(* IEC 61131-3 sources: daoli-st-library/DL_Algo (part 10) *)

(* ---- FB_DL_CoolingTowerApproachCalc.st ---- *)
//==============================================================================
// 功能块：FB_DL_CoolingTowerApproachCalc ｜ 中文名称：冷却塔逼近度计算与风机台数优化建议
// 所属子库：DL_Algo ｜ 版本：v1.0.0 ｜ 兼容：CODESYS V3.5+ / TwinCAT 3 / 汇川 InoProShop
// 功能描述：逼近度 = 冷却水出水温度 − 湿球温度（湿球由
//           FC_DL_WetBulbTempCalc v1.1.0 计算，组合调用不内联）；逼近度
//           滑动均值（1~60 拍窗）进入目标带判断；带外给出增/减风机台数
//           建议（单拍脉冲），带内保持。优化纪律：逼近度优先、N+1 冗余
//           （减台不低于 1 台）、换台最小间隔（tMinStageTime，被阻延沿
//           发一次 3402 提示）、湿球贴物理极限逼近度时加机无益（禁止
//           建议加机）。只出建议，不直接控风机（启停时序由上位轮值件
//           裁决，本件零执行输出）。
// 开源溯源 (Origin)：道莅原创实现（参考 公开工程惯例 分类与参数域）
// 单位表：温度[摄氏度] / 相对湿度[%] / 大气压[Pa] / 逼近度[K] / 台数[台] / 换台间隔[min] / 均值窗[拍]
// 错误码表：16#0002_3401 信息级（逼近度小于 0，出水低于湿球，传感器可疑，
//           不给任何换台建议，不置 bError）/ 16#0002_3402 信息级（换台
//           请求被最小间隔阻延，阻延沿发一次，不置 bError）/
//           16#0002_3405 预留禁用（不得挪用）/ 16#0002_3410 故障级（台
//           数或算法组态非法，置 bError）/ 16#0002_3411 故障级（输入非
//           有限或湿球件故障透传，置 bError）/ 16#0002_3412 预留禁用
//           （不得挪用）
// 状态机：E_DL_ApproachState（eIdle=0 / eWarmup=10 / eMonitor=20 /
//           eStageUpPending=30 / eStageDownPending=40 / eFault=99），
//           CASE 含 ELSE 兜底，ELSE 复用 3411（§3 未为本件单列兜底槽，
//           不得越段加码）并回 eFault、脉冲全撤、建议保持（安全侧）
// 边界行为：① 湿球件 bError 或 bValid 为假 → 透传为故障 3411 +
//           bWetBulbFault，锁存型标志只在故障相处置（R115），下游信息级
//           码（钳位提示）不升格；② fApproachK 小于 0（热力学不可能，
//           传感器可疑）→ 信息 3401 + bValid := FALSE + 不给任何换台
//           建议，可疑样本不入均值窗（防污染统计）；③ nFanRunning 大于
//           nFanTotal 或 nFanTotal 小于 1 或均值窗/目标/带宽组态非法 →
//           故障 3410；④ 浮点输入非有限 → 故障 3411；⑤ 换台请求受
//           tMinStageTime 约束，被阻延 → 信息 3402（阻延沿发一次，不每
//           拍刷），阻延期间挂 eStageUpPending/eStageDownPending，退出
//           条件两条：间隔到且需求仍在（发请求回 eMonitor）或带偏差
//           消失/需求翻转（不发请求回 eMonitor）；⑥ 湿球贴物理极限逼
//           近度（常量 2.0 K）且台数已满 → bNoFurtherGain，禁止建议加
//           机；首次换台请求不受守卫约束（上电无历史换台）；⑦ 失能 →
//           建议台数保持、脉冲全撤、bValid := FALSE；⑧ 恢复首拍窗口
//           清空重走暖机；守卫定时器经请求签发「断输入一拍」重启计时
//           （R40 家族）；⑨ 上电首拍 bValid := FALSE。
// 修订历史：v1.0.0 2026-11-17 首版（R25 派单 · §4.3）
//==============================================================================
(*------------------------------------------------------------------------------
 * 枚举: E_DL_ApproachState（归属 DL_Algo，与 FB_DL_CoolingTowerApproachCalc 同文件）
 *----------------------------------------------------------------------------*)
TYPE E_DL_ApproachState :
(
    eIdle             := 0,   // 失能/待机：建议保持，脉冲全撤 / Idle: suggestion held, pulses withdrawn
    eWarmup           := 10,  // 暖机：均值窗未满，只观测不出建议 / Warmup: window not full, observe only
    eMonitor          := 20,  // 监视：带内保持或按需即时发换台请求 / Monitor: hold in band or issue request at once
    eStageUpPending   := 30,  // 增台请求被最小间隔阻延，等守卫计时 / Increase request blocked by min interval
    eStageDownPending := 40,  // 减台请求被最小间隔阻延，等守卫计时 / Decrease request blocked by min interval
    eFault            := 99   // 故障兜底态：组态非法/非有限/下游透传 / Fault fallback
);
END_TYPE
FUNCTION_BLOCK FB_DL_CoolingTowerApproachCalc
VAR_INPUT
    fCondOutC        : LREAL;                  // 冷却水出水温度 [摄氏度] / Condenser water outlet temperature [degC]
    fAmbDryC         : LREAL;                  // 环境干球温度 [摄氏度] / Ambient dry-bulb temperature [degC]
    fRhPct           : LREAL;                  // 环境相对湿度 [百分数] / Ambient relative humidity [percent]
    fPressPa         : LREAL := 101325.0;      // 大气压 [Pa]，引脚注入非魔法数 / Atmospheric pressure [Pa], pin-injected
    nFanTotal        : INT;                    // 可投风机台数 [台]，1~8 / Total available fans, 1~8
    nFanRunning      : INT;                    // 当前运行台数 [台]，0~8 / Currently running fans, 0~8
    fApproachTargetK : LREAL := 4.0;           // 目标逼近度 [K] / Target approach [K]
    fApproachTolK    : LREAL := 0.5;           // 逼近度带宽半宽 [K] / Approach band half-width [K]
    tMinStageTime    : TIME := T#5M;           // 换台最小间隔 [min] / Minimum interval between stage changes [min]
    nWinSamples      : INT := 10;              // 均值窗长度 [拍]，1~60 / Moving-average window length, 1~60
    bEnable          : BOOL;                   // 总使能 / Master enable
    bReset           : BOOL;                   // 复位，上升沿清状态与窗口 / Reset, rising edge clears state and window
END_VAR
VAR_OUTPUT
    fWetBulbC        : LREAL;                  // 湿球温度 [摄氏度]，下游件输出透传 / Wet-bulb temperature [degC], passed through
    fApproachK       : LREAL;                  // 即时逼近度 [K]，出水减湿球 / Instantaneous approach [K]
    fApproachAvgK    : LREAL;                  // 逼近度滑动均值 [K] / Moving-average approach [K]
    nFanCmd          : INT;                    // 建议运行台数 [台]，失能保持 / Suggested running fans, held on disable
    bIncReq          : BOOL;                   // 增台建议，单拍脉冲 / Increase suggestion, one-scan pulse
    bDecReq          : BOOL;                   // 减台建议，单拍脉冲 / Decrease suggestion, one-scan pulse
    bNoFurtherGain   : BOOL;                   // 湿球已贴物理极限逼近度，加机无益 / Wet bulb at physical floor, more fans useless
    bWetBulbFault    : BOOL;                   // 湿球下游件故障透传标志，只在故障相处置 / Wet-bulb downstream fault pass-through flag
    eErr             : UDINT;                  // 错误码，0 = 无错，码位 16#0002_3401 起信息级、16#0002_3410 起故障级（分带见错误码表） / Error code, 0 = no error, band info/fault per the code table
    bError           : BOOL;                   // 故障级标志，仅故障级错误置位 / Fault-class flag, set only on fault-level codes
    bValid           : BOOL;                   // 建议数据可用标志，失能/故障闸显式 FALSE / Suggestion usable flag, explicit FALSE on disable/fault gates
    eState           : E_DL_ApproachState;     // 主状态机当前状态 / Current state of the main state machine
END_VAR
VAR
    fWbOut           : LREAL;                  // 湿球件输出暂存 [摄氏度] / Wet-bulb output staging [degC]
    bWbClamped       : BOOL;                   // 湿球件钳位标志透传 / Wet-bulb clamped flag pass-through
    eWbErr           : UDINT;                  // 湿球件错误码暂存 / Wet-bulb error code staging
    bWbErr           : BOOL;                   // 湿球件故障标志暂存 / Wet-bulb fault flag staging
    bWbOk            : BOOL;                   // 湿球件可用且无故障 / Wet-bulb usable and fault-free
    fbReset          : R_TRIG;                 // 复位上升沿检测实例 / Reset rising edge detector
    fbBlockTrig      : R_TRIG;                 // 换台阻延上升沿检测实例（3402 一次触发）/ Stage-block rising edge detector, 3402 once per edge
    fbStageGuard     : TON;                    // 换台最小间隔守卫定时器 / Stage interval guard timer
    bGuardKick       : BOOL;                   // 守卫定时器断输入一拍标志（R40 家族）/ Guard timer one-scan kick flag
    afWinBuf         : ARRAY[0..59] OF LREAL;  // 逼近度滑动窗缓冲 [K] / Approach sliding window buffer [K]
    nWinIdx          : INT;                    // 窗写指针 [—] / Window write pointer
    uWinFill         : UDINT;                  // 窗已填充数 [拍] / Window filled count
    fWinSum          : LREAL;                  // 窗内累加和 [K]，增量维护 / Window running sum [K], incrementally maintained
    fApproachNew     : LREAL;                  // 本拍新逼近度样本 [K] / New approach sample this scan [K]
    bBadSensor       : BOOL;                   // 逼近度小于 0，传感器可疑 / Approach negative, sensor suspect
    bNeedInc         : BOOL;                   // 本拍需要增台（实时重算）/ Increase needed this scan, recomputed
    bNeedDec         : BOOL;                   // 本拍需要减台（实时重算）/ Decrease needed this scan, recomputed
    bGuardOk         : BOOL;                   // 守卫放行：无历史换台或间隔已满 / Guard released: no history or interval elapsed
    bBlockedNow      : BOOL;                   // 本拍换台请求被阻延 / Stage request blocked this scan
    bStageEverReq    : BOOL;                   // 激活以来是否签发过换台请求 / Any stage request issued since activation
    bFanCmdInit      : BOOL;                   // 建议台数是否已初始化 / Suggestion count initialized flag
    bActiveCalc      : BOOL;                   // 本拍处于可计算状态（暖机/监视/阻延挂起）/ Computable state this scan
END_VAR
VAR CONSTANT
    DL_CTWR_CODE_INFO_1 : UDINT := 16#0002_3401;   // 信息级槽 1（逼近度小于 0） / info slot 1
    DL_CTWR_CODE_INFO_2 : UDINT := 16#0002_3402;   // 信息级槽 2（换台请求被阻延） / info slot 2
    DL_CTWR_CODE_RSV_1  : UDINT := 16#0002_3405;   // 预留禁用（不得挪用） / reserved, do not use
    DL_CTWR_CODE_FLT_1  : UDINT := 16#0002_3410;   // 故障级槽 1（台数或组态非法） / fault slot 1
    DL_CTWR_CODE_FLT_2  : UDINT := 16#0002_3411;   // 故障级槽 2（非有限或湿球透传） / fault slot 2
    DL_CTWR_CODE_RSV_2  : UDINT := 16#0002_3412;   // 预留禁用（不得挪用） / reserved, do not use
    DL_AP_ZERO       : LREAL := 0.0;           // 零值常量，避免裸字面量 [—] / Zero constant, avoids a bare literal
    DL_AP_INF        : LREAL := 1.7976931348623157E308;  // LREAL 幅值上限，Inf 判据 / LREAL magnitude ceiling, Inf criterion
    DL_AP_TOL        : LREAL := 1.0E-6;        // 浮点比较容差 [—] / Float comparison tolerance
    DL_AP_WIN_MAX    : INT   := 60;            // 均值窗长度上限 [拍] / Moving-average window ceiling
    DL_AP_FAN_MAX    : INT   := 8;             // 风机台数上限 [台] / Fan count ceiling
    DL_AP_FAN_MIN    : INT   := 1;             // N+1 冗余最低运行台数 [台] / Minimum running fans for N+1 redundancy
    DL_AP_PHYS_FLOOR : LREAL := 2.0;           // 物理极限逼近度 [K]，贴限判加机无益 / Physical floor approach [K], gain-limit criterion
END_VAR

(*------------------------------------------------------------------------------
 * 段 1｜无条件刷新区（红线 5）：沿检测与守卫定时器在任何分支之外周期调用
 *----------------------------------------------------------------------------*)
fbReset(CLK := bReset);                        // 复位沿检测无条件刷新 / reset edge refreshed unconditionally
fbStageGuard(IN := bEnable AND NOT bGuardKick, // 断输入一拍重启计时（R40 家族）/ break input one scan to restart timing
             PT := tMinStageTime);             // 守卫门槛 = 换台最小间隔 / guard threshold = min stage interval
bGuardKick := FALSE;                           // kick 标志单拍自清（本拍签发请求时由状态机重置位）/ kick flag self-clears, state machine re-sets on issue

(*------------------------------------------------------------------------------
 * 段 2｜复位沿处理（改写置于沿后，防吞沿 R39）
 *----------------------------------------------------------------------------*)
IF fbReset.Q THEN
    eState        := E_DL_ApproachState.eIdle;
    eErr          := 16#0000_0000;             // 复位清码 / reset clears code
    bError        := FALSE;                    // 复位清故障 / reset clears fault
    uWinFill      := 0;                        // 窗口清空重走暖机 / window cleared, warmup again
    nWinIdx       := 0;                        // 写指针归零 / write pointer zeroed
    fWinSum       := DL_AP_ZERO;               // 累加和清零 / sum zeroed
    fApproachAvgK := DL_AP_ZERO;               // 均值出口清零 / average output zeroed
    bIncReq       := FALSE;                    // 脉冲全撤 / pulses withdrawn
    bDecReq       := FALSE;                    // 脉冲全撤 / pulses withdrawn
    bNoFurtherGain := FALSE;                   // 贴限标志清除 / gain-limit flag cleared
    bBadSensor    := FALSE;                    // 传感器可疑标志清除 / suspect flag cleared
    bStageEverReq := FALSE;                    // 换台历史清零，首个请求放行 / stage history cleared, first request released
    bFanCmdInit   := FALSE;                    // 建议台数待重初始化 / suggestion count re-initialized
END_IF

(*------------------------------------------------------------------------------
 * 段 3｜非有限输入闸（浮点引脚逐个：NaN 自反判 + Inf 幅值上限判，R79）
 *----------------------------------------------------------------------------*)
IF (fCondOutC <> fCondOutC) OR (ABS(fCondOutC) >= DL_AP_INF)
   OR (fAmbDryC <> fAmbDryC) OR (ABS(fAmbDryC) >= DL_AP_INF)
   OR (fRhPct <> fRhPct) OR (ABS(fRhPct) >= DL_AP_INF)
   OR (fPressPa <> fPressPa) OR (ABS(fPressPa) >= DL_AP_INF)
   OR (fApproachTargetK <> fApproachTargetK) OR (ABS(fApproachTargetK) >= DL_AP_INF)
   OR (fApproachTolK <> fApproachTolK) OR (ABS(fApproachTolK) >= DL_AP_INF) THEN
    eState := E_DL_ApproachState.eFault;
    eErr   := DL_CTWR_CODE_FLT_2;                  // 故障级：输入非有限 / fault: non-finite input
    bError := TRUE;                            // 故障级必置 bError（R45 配对）/ fault-class pairs with bError
    bValid := FALSE;                           // 输出不可用 / outputs unusable
    bIncReq := FALSE;                          // 脉冲全撤安全侧 / pulses withdrawn, safe side
    bDecReq := FALSE;                          // 脉冲全撤安全侧 / pulses withdrawn, safe side
    bNoFurtherGain := FALSE;                   // 故障态不判贴限 / gain-limit not judged in fault
    RETURN;
END_IF

(*------------------------------------------------------------------------------
 * 段 4｜组态合法性闸（台数域/主从关系/窗长/目标/带宽）
 *----------------------------------------------------------------------------*)
IF (nFanTotal < DL_AP_FAN_MIN) OR (nFanTotal > DL_AP_FAN_MAX)
   OR (nFanRunning < 0) OR (nFanRunning > nFanTotal)
   OR (nWinSamples < 1) OR (nWinSamples > DL_AP_WIN_MAX)
   OR (fApproachTargetK <= DL_AP_TOL) OR (fApproachTolK <= DL_AP_TOL) THEN
    eState := E_DL_ApproachState.eFault;
    eErr   := DL_CTWR_CODE_FLT_1;                  // 故障级：台数或算法组态非法 / fault: fan or algorithm config invalid
    bError := TRUE;                            // 故障级必置 bError（R45 配对）/ fault-class pairs with bError
    bValid := FALSE;                           // 输出不可用 / outputs unusable
    bIncReq := FALSE;                          // 脉冲全撤安全侧 / pulses withdrawn, safe side
    bDecReq := FALSE;                          // 脉冲全撤安全侧 / pulses withdrawn, safe side
    bNoFurtherGain := FALSE;                   // 故障态不判贴限 / gain-limit not judged in fault
    RETURN;
END_IF

(*------------------------------------------------------------------------------
 * 段 5｜湿球组合调用：每拍恰好一次，不内联不复制（R115 透传纪律）
 *----------------------------------------------------------------------------*)
FC_DL_WetBulbTempCalc(fTempC := fAmbDryC, fRh := fRhPct, fPress := fPressPa,
                      fWetBulbC => fWbOut, bClamped => bWbClamped,
                      eErr => eWbErr, bError => bWbErr, bValid => bWbOk);
fWetBulbC := fWbOut;                           // 湿球出口透传 / wet-bulb output pass-through
IF bWbErr OR (NOT bWbOk) THEN
    bWetBulbFault := TRUE;                     // 下游故障透传标志 / downstream fault pass-through flag
ELSE
    bWetBulbFault := FALSE;                    // 下游正常，信息级钳位不升格 / downstream ok, info-level clamp not escalated
END_IF

(*------------------------------------------------------------------------------
 * 段 6｜逼近度计算与滑动窗维护（仅在使能、湿球可用、传感器不可疑时推进）
 *----------------------------------------------------------------------------*)
bActiveCalc := bEnable AND (NOT bWetBulbFault)
           AND (eState = E_DL_ApproachState.eWarmup
             OR eState = E_DL_ApproachState.eMonitor
             OR eState = E_DL_ApproachState.eStageUpPending
             OR eState = E_DL_ApproachState.eStageDownPending);  // 可计算状态判据 / computable-state predicate
bBadSensor := FALSE;                           // 传感器可疑标志逐拍重判 / suspect flag re-judged per scan
IF bActiveCalc THEN
    fApproachK := fCondOutC - fWetBulbC;       // 即时逼近度 = 出水 − 湿球 [K] / instantaneous approach = outlet minus wet bulb
    bBadSensor := fApproachK < -DL_AP_TOL;     // 热力学不可能，传感器可疑 / thermodynamically impossible, sensor suspect
    IF bBadSensor THEN
        // 可疑样本不入窗，均值保持（防污染统计）/ suspect sample not pushed, average held
    ELSE
        IF uWinFill < INT_TO_UDINT(nWinSamples) THEN
            uWinFill := uWinFill + 1;          // 窗未满：填充数递增 / window not full: fill count up
            fWinSum := fWinSum + fApproachK;   // 累加和并入新样本 / sum absorbs new sample
            afWinBuf[nWinIdx] := fApproachK;   // 写入当前槽 / write current slot
        ELSE
            fWinSum := fWinSum - afWinBuf[nWinIdx] + fApproachK;  // 窗满：换出旧值并入新值 / window full: swap out old, absorb new
            afWinBuf[nWinIdx] := fApproachK;   // 覆盖当前槽 / overwrite current slot
        END_IF
        nWinIdx := (nWinIdx + 1) MOD nWinSamples;  // 写指针环形推进，nWinSamples 已闸大于 0 / ring-advance write pointer, divisor gated
        fApproachAvgK := fWinSum / UDINT_TO_LREAL(uWinFill);  // 均值 = 和/填充数，填充数已闸大于 0 / average, fill count gated
    END_IF
END_IF

(*------------------------------------------------------------------------------
 * 段 7｜决策块：带偏差实时重算（阻延挂起态也用同一决策，需求翻转即退出）
 *----------------------------------------------------------------------------*)
bNeedInc := FALSE;                             // 增台需求逐拍重判 / increase need re-judged per scan
bNeedDec := FALSE;                             // 减台需求逐拍重判 / decrease need re-judged per scan
bNoFurtherGain := FALSE;                       // 贴限标志逐拍重判，非计算态不残留 / gain-limit flag re-judged per scan
bGuardOk := (NOT bStageEverReq) OR fbStageGuard.Q;  // 守卫放行：无历史换台或最小间隔已满 / guard released
IF bActiveCalc AND (NOT bBadSensor) THEN
    IF NOT bFanCmdInit THEN
        nFanCmd := nFanRunning;                // 建议台数首拍初始化为当前运行台数 / suggestion initialized to running count
        bFanCmdInit := TRUE;                   // 初始化完成 / initialization done
    END_IF
    bNoFurtherGain := (fApproachK <= DL_AP_PHYS_FLOOR) AND (nFanRunning >= nFanTotal);  // 贴物理极限且台数已满，加机无益 / at physical floor with all fans on
    IF (fApproachAvgK - fApproachTargetK) > fApproachTolK THEN
        bNeedInc := (nFanRunning < nFanTotal) AND (NOT bNoFurtherGain);  // 偏热且有余量：增台 / too hot with headroom: increase
    ELSIF (fApproachTargetK - fApproachAvgK) > fApproachTolK THEN
        bNeedDec := (nFanRunning > DL_AP_FAN_MIN);  // 偏冷且高于冗余下限：减台 / too cold above redundancy floor: decrease
    END_IF
END_IF

(*------------------------------------------------------------------------------
 * 段 8｜阻延沿检测（无条件周期调用，CLK 为本拍阻延判据，3402 沿发一次）
 *----------------------------------------------------------------------------*)
bBlockedNow := bActiveCalc AND (NOT bBadSensor) AND (bNeedInc OR bNeedDec) AND (NOT bGuardOk);  // 本拍阻延判据 / blocked predicate this scan
fbBlockTrig(CLK := bBlockedNow);               // 阻延沿检测无条件刷新 / block edge refreshed unconditionally

(*------------------------------------------------------------------------------
 * 段 9｜状态机：CASE 含 ELSE 兜底。bIncReq/bDecReq 为单拍脉冲：本段开头
 *       先无条件撤脉冲，状态机内按需重置位（先撤后置，不跨拍残留）。
 *----------------------------------------------------------------------------*)
bIncReq := FALSE;                              // 单拍脉冲先撤 / one-scan pulse withdrawn first
bDecReq := FALSE;                              // 单拍脉冲先撤 / one-scan pulse withdrawn first

CASE eState OF

    E_DL_ApproachState.eIdle:
        bValid := FALSE;                       // 失能闸显式不可用（R72）/ explicit FALSE on disable gate
        eErr := 16#0000_0000;                  // 待机无错 / no error in idle
        bError := FALSE;                       // 待机无故障 / no fault in idle
        bWetBulbFault := FALSE;                // 待机不透传故障相（R115：只在故障相处置）/ pass-through only in fault phase
        bNoFurtherGain := FALSE;               // 待机不判贴限 / gain-limit not judged in idle
        IF bEnable THEN
            IF bWetBulbFault THEN
                eState := E_DL_ApproachState.eFault;   // 湿球不可用直接进故障 / unusable wet bulb enters fault
                eErr := DL_CTWR_CODE_FLT_2;    // 故障级：湿球件故障透传 / fault: wet-bulb pass-through
                bError := TRUE;                // 故障级必置 bError / fault-class pairs with bError
            ELSE
                eState := E_DL_ApproachState.eWarmup;  // 使能且湿球可用进暖机 / enable with valid wet bulb enters warmup
            END_IF
        END_IF

    E_DL_ApproachState.eWarmup:
        eErr := 16#0000_0000;                  // 暖机默认无错 / warmup defaults to no error
        bError := FALSE;                       // 暖机默认无故障 / warmup defaults to no fault
        bValid := FALSE;                       // 暖机期窗口未满不可用 / unusable during warmup
        IF NOT bEnable THEN
            eState := E_DL_ApproachState.eIdle;        // 失能回待机 / disable returns to idle
        ELSIF bWetBulbFault THEN
            eState := E_DL_ApproachState.eFault;       // 下游故障进故障态 / downstream fault enters fault state
            eErr := DL_CTWR_CODE_FLT_2;        // 故障级：湿球件故障透传 / fault: wet-bulb pass-through
            bError := TRUE;                    // 故障级必置 bError / fault-class pairs with bError
        ELSIF bBadSensor THEN
            eErr := DL_CTWR_CODE_INFO_1;       // 信息级：逼近度小于 0，传感器可疑 / info: negative approach, sensor suspect
            bValid := FALSE;                   // 传感器可疑，不给建议 / suspect sensor, no advice
        ELSIF uWinFill >= INT_TO_UDINT(nWinSamples) THEN
            eState := E_DL_ApproachState.eMonitor;     // 均值窗已满进监视 / window full enters monitor
        END_IF

    E_DL_ApproachState.eMonitor:
        IF NOT bEnable THEN
            eState := E_DL_ApproachState.eIdle;        // 失能回待机 / disable returns to idle
            bValid := FALSE;                   // 失能闸显式不可用（R72）/ explicit FALSE on disable gate
        ELSIF bWetBulbFault THEN
            eState := E_DL_ApproachState.eFault;
            eErr := DL_CTWR_CODE_FLT_2;        // 故障级：湿球件故障透传 / fault: wet-bulb pass-through
            bError := TRUE;                    // 故障级必置 bError / fault-class pairs with bError
            bValid := FALSE;                   // 故障闸显式不可用 / explicit FALSE on fault gate
        ELSIF bBadSensor THEN
            eErr := DL_CTWR_CODE_INFO_1;       // 信息级：逼近度小于 0 / info: negative approach
            bError := FALSE;                   // 信息级不置 bError / info never raises bError
            bValid := FALSE;                   // 传感器可疑，不给建议（边界行为②）/ suspect sensor, no advice
        ELSE
            eErr := 16#0000_0000;              // 正常监视清码 / normal monitor clears code
            bError := FALSE;                   // 正常监视清故障 / normal monitor clears fault
            bValid := TRUE;                    // 建议数据可用 / suggestion usable
            IF bNeedInc OR bNeedDec THEN
                IF bGuardOk THEN
                    IF bNeedInc THEN
                        bIncReq := TRUE;       // 增台建议单拍脉冲 / increase pulse
                        nFanCmd := nFanRunning + 1;    // 建议台数加一 / suggested count up
                    ELSE
                        bDecReq := TRUE;       // 减台建议单拍脉冲 / decrease pulse
                        nFanCmd := nFanRunning - 1;    // 建议台数减一 / suggested count down
                    END_IF
                    bStageEverReq := TRUE;     // 记录换台历史 / record stage history
                    bGuardKick := TRUE;        // 守卫定时器断输入一拍重启 / guard timer kicked one scan
                ELSE
                    IF bNeedInc THEN
                        eState := E_DL_ApproachState.eStageUpPending;  // 增台请求被阻延挂起 / increase request blocked, pending
                    ELSE
                        eState := E_DL_ApproachState.eStageDownPending;  // 减台请求被阻延挂起 / decrease request blocked, pending
                    END_IF
                END_IF
            END_IF
        END_IF

    E_DL_ApproachState.eStageUpPending:
        IF NOT bEnable THEN
            eState := E_DL_ApproachState.eIdle;
            bValid := FALSE;                   // 失能闸显式不可用（R72）/ explicit FALSE on disable gate
        ELSIF bWetBulbFault THEN
            eState := E_DL_ApproachState.eFault;
            eErr := DL_CTWR_CODE_FLT_2;
            bError := TRUE;
            bValid := FALSE;
        ELSIF bBadSensor THEN
            eState := E_DL_ApproachState.eMonitor;     // 传感器可疑，需求作废回监视 / suspect sensor, need voided, back to monitor
            eErr := DL_CTWR_CODE_INFO_1;
            bError := FALSE;
            bValid := FALSE;
        ELSIF NOT bNeedInc THEN
            eState := E_DL_ApproachState.eMonitor;     // 需求消失退出（第二条退出条件）/ need vanished, second exit condition
            eErr := 16#0000_0000;              // 回监视清码 / clear code on return
            bValid := TRUE;                    // 回监视数据可用 / usable on return
        ELSIF fbStageGuard.Q THEN
            bIncReq := TRUE;                   // 间隔到且需求仍在：签发增台 / interval elapsed with need: issue increase
            nFanCmd := nFanRunning + 1;        // 建议台数加一 / suggested count up
            bStageEverReq := TRUE;             // 记录换台历史 / record stage history
            bGuardKick := TRUE;                // 守卫定时器断输入一拍重启 / guard timer kicked one scan
            eState := E_DL_ApproachState.eMonitor;     // 签发后回监视 / back to monitor after issue
            eErr := 16#0000_0000;              // 阻延解除清码 / clear code on release
            bValid := TRUE;                    // 数据可用 / usable
        ELSE
            bValid := TRUE;                    // 挂起期间建议数据仍可用 / suggestion usable while pending
        END_IF

    E_DL_ApproachState.eStageDownPending:
        IF NOT bEnable THEN
            eState := E_DL_ApproachState.eIdle;
            bValid := FALSE;                   // 失能闸显式不可用（R72）/ explicit FALSE on disable gate
        ELSIF bWetBulbFault THEN
            eState := E_DL_ApproachState.eFault;
            eErr := DL_CTWR_CODE_FLT_2;
            bError := TRUE;
            bValid := FALSE;
        ELSIF bBadSensor THEN
            eState := E_DL_ApproachState.eMonitor;     // 传感器可疑，需求作废回监视 / suspect sensor, need voided, back to monitor
            eErr := DL_CTWR_CODE_INFO_1;
            bError := FALSE;
            bValid := FALSE;
        ELSIF NOT bNeedDec THEN
            eState := E_DL_ApproachState.eMonitor;     // 需求消失退出（第二条退出条件）/ need vanished, second exit condition
            eErr := 16#0000_0000;              // 回监视清码 / clear code on return
            bValid := TRUE;                    // 回监视数据可用 / usable on return
        ELSIF fbStageGuard.Q THEN
            bDecReq := TRUE;                   // 间隔到且需求仍在：签发减台 / interval elapsed with need: issue decrease
            nFanCmd := nFanRunning - 1;        // 建议台数减一 / suggested count down
            bStageEverReq := TRUE;             // 记录换台历史 / record stage history
            bGuardKick := TRUE;                // 守卫定时器断输入一拍重启 / guard timer kicked one scan
            eState := E_DL_ApproachState.eMonitor;     // 签发后回监视 / back to monitor after issue
            eErr := 16#0000_0000;              // 阻延解除清码 / clear code on release
            bValid := TRUE;                    // 数据可用 / usable
        ELSE
            bValid := TRUE;                    // 挂起期间建议数据仍可用 / suggestion usable while pending
        END_IF

    ELSE
        eState := E_DL_ApproachState.eFault;   // 非法状态兜底 / illegal-state fallback
        eErr   := DL_CTWR_CODE_FLT_2;          // 兜底复用故障级槽 2（§3 未单列兜底槽，不得越段加码）/ fallback reuses fault slot 2
        bError := TRUE;                        // 故障级必置 bError / fault-class pairs with bError
        bValid := FALSE;                       // 输出不可用 / outputs unusable
        bIncReq := FALSE;                      // 脉冲全撤安全侧 / pulses withdrawn, safe side
        bDecReq := FALSE;                      // 脉冲全撤安全侧 / pulses withdrawn, safe side
END_CASE

(*------------------------------------------------------------------------------
 * 段 10｜信息级收口：阻延沿发一次 3402（不每拍刷，见边界行为⑤）
 *----------------------------------------------------------------------------*)
IF fbBlockTrig.Q THEN
    eErr := DL_CTWR_CODE_INFO_2;               // 信息级：换台请求被最小间隔阻延 / info: stage request blocked by interval
    bError := FALSE;                           // 信息级不置 bError / info never raises bError
END_IF
END_FUNCTION_BLOCK

(* ---- FB_DL_CoolingTowerOpt.st ---- *)
(*
  Component : FB_DL_CoolingTowerOpt
  Category  : DL_Algo
  Type      : FB
  Version   : 1.0.0
  CodeSeg   : 16#02_3_5F
  Summary   : 冷却塔群控逼近度优化：湿球逼近度控制律 + 塔群投切决策（最小开机数 + 防震荡死区）。
              Cooling tower approach optimization: wet-bulb approach control law plus staging with min-on units and deadband.
  溯源声明  : 道莅自研 clean-room
  边界安全  : 温度/台数非有限（NaN 自反 + Inf 上限）拦截；塔数域闸（1..8，防数组越界）；
              最小开机数域闸（1..nTowers，防全停）与投切错峰窗（自复位 TON）防频繁投切；
              投切决策带对称死区（防震荡）；风机设定值输出过 RateLimiter 限速；
              全浮点比较带 fEps 容差；计数防回卷。
  复用      : 无
*)

FUNCTION_BLOCK FB_DL_CoolingTowerOpt
VAR_INPUT
    bRun          : BOOL;              (* 优化使能 · Enable *)
    fWetBulbC     : LREAL;             (* 湿球温度 [degC] · Wet-bulb temperature *)
    fOutTC        : LREAL;             (* 塔群出水温度 [degC] · Tower outlet temperature *)
    fApprTargetC  : LREAL := 3.0;      (* 逼近度目标 [K] · Approach target *)
    fDeadK        : LREAL := 0.5;      (* 投切死区 [K]，防震荡 · Staging deadband *)
    nTowersAvail  : INT   := 4;        (* 可用塔数 [台]，域 1 到 8 · Available towers *)
    nMinOn        : INT   := 1;        (* 最小开机数 [台] · Minimum on units *)
    tStaggerMs    : TIME  := T#30000MS; (* 投切错峰窗 [ms] · Stagger window *)
    fFanStepPct   : LREAL := 2.0;      (* 风机设定每拍最大步进 [％] · Fan setpoint max step *)
    fEps          : LREAL := 1.0E-6;   (* 浮点判零容差 [实数域] · Floating zero tolerance *)
END_VAR
VAR_OUTPUT
    aTowerCmd : ARRAY[1..8] OF BOOL;    (* 各塔投切指令 [引脚] · Per-tower commands *)
    nRunCnt   : INT;                    (* 当前开机数 [台] · Currently running count *)
    fApprNowC : LREAL;                  (* 当前逼近度 [K] · Current approach *)
    fFanSetPct: LREAL;                  (* 风机群设定值输出 [％]，已限速 · Rate-limited fan setpoint *)
    bError    : BOOL;                   (* 故障标志，与故障码配对 · Fault flag paired with codes *)
    uErrorId  : UDINT;                  (* 事件码 16#0000_005F，0 无事件 · Event code *)
END_VAR
VAR
    _eState   : (eStHold := 0, eStAdd := 1, eStDrop := 2);  (* 内部决策状态 / Internal decision state *)
    uCode     : WORD;    (* 码位暂存，每拍重算 [码] · Code staging *)
    tonStagger: TON;     (* 投切错峰窗 [ms]，自复位振荡 · Stagger timer, self-reset *)
    bSigOk    : BOOL;    (* 输入有效标志 · Input validity flag *)
    bTick     : BOOL;    (* 错峰窗到点脉冲 [脉冲] · Stagger tick pulse *)
    nI        : INT;     (* 塔循环下标 [索引] · Tower loop index *)
    fFanTgt   : LREAL;   (* 风机设定目标 [％] · Fan setpoint target *)
    fStep     : LREAL;   (* 本拍设定步进 [％] · Actual step this scan *)
    nCycles   : UDINT;   (* 有效拍计数 [拍]，防回卷 · Valid scan count *)
END_VAR
VAR CONSTANT
    DL_CTO_NMAX  : INT   := 8;          (* 塔数上限 [台]，与数组一致 · Tower cap *)
    DL_CTO_FANHI : LREAL := 100.0;      (* 风机设定上限 [％] · Fan setpoint cap high *)
    DL_CTO_FANLO : LREAL := 40.0;       (* 风机设定下限 [％] · Fan setpoint cap low *)
    DL_CTO_WRAP  : UDINT := 4294967290; (* 计数防回卷余量 [拍] · Counter wrap guard *)
END_VAR

(* === 段 0 · 实例刷新（每拍无条件，红线 7）=== *)
tonStagger(IN := NOT tonStagger.Q, PT := tStaggerMs);   (* 错峰窗自复位振荡 / Self-reset stagger window *)
bTick := tonStagger.Q;                                  (* 窗到点脉冲 / Stagger tick *)

(* === 段 1 · 输入校验与量程闸 === *)
uCode := 16#0000;                       // 每拍清码（可达清零基线）/ Clear codes each scan
bSigOk := (fWetBulbC = fWetBulbC) AND (fOutTC = fOutTC)             // 非有限拦截 / Non-finite guard
          AND (ABS(fWetBulbC) < 1.0E308) AND (ABS(fOutTC) < 1.0E308) // Inf 上限判据 / Inf limit
          AND (nTowersAvail >= 1) AND (nTowersAvail <= DL_CTO_NMAX)  // 塔数域闸，防越界 / Tower count gate
          AND (nMinOn >= 1) AND (nMinOn <= nTowersAvail)             // 最小开机数域闸，防全停 / Min-on gate
          AND (fDeadK >= 0.0) AND (fFanStepPct > 0.0);               // 死区/步进域闸 / Deadband and step gates
IF NOT bSigOk THEN
    uCode := 16#005F;                   // 故障级：域外，决策冻结 / Fault: domain invalid
END_IF

(* === 段 2 · 主逻辑：逼近度控制律与投切决策 === *)
IF bSigOk THEN
    fApprNowC := fOutTC - fWetBulbC;    (* 当前逼近度 [K] / Current approach *)
    IF NOT bRun THEN
        _eState := eStHold;             (* 撤使决策保持 / Hold on disable *)
        FOR nI := 1 TO DL_CTO_NMAX DO
            aTowerCmd[nI] := FALSE;     (* 撤使全停 / All off on disable *)
        END_FOR
        nRunCnt := 0;                   (* 开机数清零 / Clear the count *)
        fFanTgt := DL_CTO_FANLO;        (* 撤使风机回下限 / Fan to low cap *)
    ELSE
        (* 决策状态机：死区外才进投切相，错峰窗内每窗一台 / One unit per window outside the deadband *)
        IF NOT bTick THEN
            _eState := eStHold;         (* 窗内保持 / Hold inside the window *)
        ELSIF fApprNowC > (fApprTargetC + fDeadK) THEN
            _eState := eStAdd;          (* 逼近度超标：投塔相 / Over target: add phase *)
        ELSIF fApprNowC < (fApprTargetC - fDeadK) THEN
            _eState := eStDrop;         (* 逼近度过低：切塔相 / Under target: drop phase *)
        ELSE
            _eState := eStHold;         (* 死区内保持（防震荡）/ Hold inside the deadband *)
        END_IF
        CASE _eState OF
            eStAdd:                     (* 投塔：找一台未开塔，保最小开机数下限之上 / Add one tower *)
                FOR nI := 1 TO nTowersAvail DO
                    IF NOT aTowerCmd[nI] THEN
                        aTowerCmd[nI] := TRUE;      (* 投入该塔 / Turn the tower on *)
                        EXIT;           (* 单台即止 / One unit only *)
                    END_IF
                END_FOR
            eStDrop:                    (* 切塔：开机数大于最小开机数才允许 / Drop only above min-on *)
                IF nRunCnt > nMinOn THEN
                    FOR nI := nTowersAvail TO 1 BY -1 DO
                        IF aTowerCmd[nI] THEN
                            aTowerCmd[nI] := FALSE; (* 切除该塔 / Turn the tower off *)
                            EXIT;       (* 单台即止 / One unit only *)
                        END_IF
                    END_FOR
                END_IF
            eStHold:                    (* 保持相：不动塔群 / Hold: no staging *)
                (* 无动作 / No action *)
        ELSE
            _eState := eStHold;         (* ELSE 兜底回保持相 / ELSE fallback to hold *)
        END_CASE
        nRunCnt := 0;                   (* 开机数重算 / Recount *)
        FOR nI := 1 TO DL_CTO_NMAX DO
            IF aTowerCmd[nI] THEN
                nRunCnt := nRunCnt + 1; (* 累加实开塔数 / Count the running towers *)
            END_IF
        END_FOR
        (* 风机设定目标：逼近度超死区升频，低于死区降频，钳上下限 / Fan target by approach *)
        IF fApprNowC > (fApprTargetC + fDeadK) THEN
            fFanTgt := fFanTgt + fFanStepPct;   (* 升频目标 / Raise target *)
        ELSIF fApprNowC < (fApprTargetC - fDeadK) THEN
            fFanTgt := fFanTgt - fFanStepPct;   (* 降频目标 / Lower target *)
        END_IF
        IF fFanTgt > DL_CTO_FANHI THEN
            fFanTgt := DL_CTO_FANHI;    (* 钳上限 / Cap high *)
        ELSIF fFanTgt < DL_CTO_FANLO THEN
            fFanTgt := DL_CTO_FANLO;    (* 钳下限 / Cap low *)
        END_IF
    END_IF
    (* RateLimiter：风机设定限速 / Rate limit the fan setpoint *)
    fStep := fFanTgt - fFanSetPct;      (* 目标差 [％] / Gap to target *)
    IF fStep > fFanStepPct THEN
        fFanSetPct := fFanSetPct + fFanStepPct;     (* 正向限速 / Positive rate limit *)
    ELSIF fStep < (-fFanStepPct) THEN
        fFanSetPct := fFanSetPct - fFanStepPct;     (* 负向限速 / Negative rate limit *)
    ELSE
        fFanSetPct := fFanTgt;          (* 一步到位 / Settle *)
    END_IF
END_IF

(* === 段 3 · 输出映射与故障码 === *)
IF bSigOk THEN
    IF nCycles < DL_CTO_WRAP THEN
        nCycles := nCycles + 1;         (* 有效拍计数 / Count valid scans *)
    END_IF
END_IF
bError := (uCode <> 16#0000);           (* 故障标志配对 / Fault flag paired *)
uErrorId := WORD_TO_UDINT(uCode);       (* 码位单点写入（16#0000_005F 形态）/ Single write point *)
END_FUNCTION_BLOCK

(* ---- FB_DL_CraneAntiSway.st ---- *)
(*
  ==================================================================
  组件名 Component  : FB_DL_CraneAntiSway
  分类   Category   : DL_Algo
  复杂度 Complexity  : 中
  版本   Version    : 1.0.0
  功能   Purpose    : 桥式起重机防摆控制。摆角/摆速反馈相位对消：补偿量
                      fCorr = K1·角度 + K2·摆速 叠加到运行速度指令；输出
                      钳位 ±fVmax；防摆-定位双模：|角度| < 角容差 且 |摆速|
                      < 速容差 时置定位带内 bInPosBand（供定位模切换判据）。
                      GitHub topics crane 线公开语义 clean-room。
  来源   Source     : T1-8-github-topics（crane 防摆公开语义）
  溯源   Origin     : 摆角/摆速相位对消为公开控制语义，clean-room 自研实现，
                      未复制任何厂商私有库源码。
  平台   Platform   : 纯 IEC 61131-3，CODESYS / TwinCAT / InoProShop 通用
  分工声明 Split     : 与 FB_DL_LookaheadVelPlanner 分工——后者做速度前瞻，
                      本件做摆动反馈补偿叠加。
  作者   Author     : 道莅代码库 · PLC 编程专家（R59）
  ------------------------------------------------------------------
  边界 Boundary     :
                      一 非有限闸（自反双判据，三输入全覆盖）：命中置 bBad
                         （本库纪律②），fVout 安全侧零；
                      二 输出硬钳位 ±fVmax 单点回夹并置 bClamped（信息级）；
                      三 失能安全语义：bEnable = FALSE 时 fVout = 0（安全侧
                         零速，防摆-定位双模声明 R191）；
                      四 补偿增益组态域由调用方保证（K1/K2 为负值使摆角正
                         馈回拉），本件不二次钳制；
                      五 无全局变量、无外部变量声明、无物理地址寻址。
  修订记录 Revision  :
    2026-11-21  v1.0.0  R59 首版（批 3 · 序号 12）
  ==================================================================
*)

FUNCTION_BLOCK FB_DL_CraneAntiSway
VAR_INPUT
    fVcmd       : LREAL := 0.0;  // 运行速度指令 [毫米每秒] / the travel velocity command [millimeter per second]
    fAngDeg     : LREAL := 0.0;  // 摆角反馈 [度] / the sway angle feedback [degree]
    fAngVelDegS : LREAL := 0.0;  // 摆速反馈 [度每秒] / the sway angular velocity feedback [degree per second]
    fK1         : LREAL := -2.0; // 摆角补偿增益 [（毫米每秒）每度] / the angle compensation gain
    fK2         : LREAL := -8.0; // 摆速补偿增益 [（毫米每秒）每（度每秒）] / the velocity compensation gain
    fVmax       : LREAL := 500.0; // 输出速度上界 [毫米每秒] / the outlet velocity bound [millimeter per second]
    fPosAngTol  : LREAL := 1.0;  // 定位带角容差 [度] / the positioning angle tolerance [degree]
    fPosVelTol  : LREAL := 2.0;  // 定位带速容差 [度每秒] / the positioning velocity tolerance [degree per second]
    bAntiSwayEn : BOOL := TRUE;  // 防摆补偿使能（定位模可关）[-] / the anti sway enable
    bEnable     : BOOL := FALSE; // 输出使能，失能安全侧零 [-] / the outlet enable, the safe zero when disabled
END_VAR
VAR_OUTPUT
    fVout     : LREAL := 0.0; // 补偿后速度输出 [毫米每秒] / the compensated velocity outlet
    fCorr     : LREAL := 0.0; // 防摆补偿量（观测用）[毫米每秒] / the anti sway compensation, observable
    bInPosBand: BOOL := FALSE; // 定位带内判据（双模切换依据）[-] / the in position band verdict
    bClamped  : BOOL := FALSE; // 输出钳位发生（信息级）[-] / the outlet clamp happened, informational
    bBad      : BOOL := FALSE; // 非有限输入实时标志 [-] / the non finite input flag
    bValid    : BOOL := FALSE; // 输出可用标志 [-] / the output usable flag
END_VAR
VAR
    _fV   : LREAL; // 补偿后速度工作量 [毫米每秒] / the compensated velocity work value
    _bFin : BOOL;  // 输入有限工作量 [-] / the input finiteness work flag
END_VAR

// 段 1｜输出预置与非有限闸（四段式，R45 + 本库纪律②）/ segment 1, the preset and the non finite gate
fVout := 0.0; // 输出预置安全零 / preset the safe zero
fCorr := 0.0; // 补偿预置零 / preset the compensation zero
bClamped := FALSE; // 钳位预置假 / preset the clamp false
bValid := FALSE; // 有效预置假 / preset the valid false
_bFin := (fVcmd = fVcmd) AND ((fVcmd - fVcmd) = (fVcmd - fVcmd)) // 指令有限 / the command finite
    AND (fAngDeg = fAngDeg) AND ((fAngDeg - fAngDeg) = (fAngDeg - fAngDeg)) // 摆角有限 / the angle finite
    AND (fAngVelDegS = fAngVelDegS) AND ((fAngVelDegS - fAngVelDegS) = (fAngVelDegS - fAngVelDegS)); // 摆速有限 / the velocity finite
bBad := NOT _bFin; // 拒收实时标志（R191 名实双出口）/ the rejection flag
IF bBad THEN // 非有限命中 / a non finite hit
    bInPosBand := FALSE; // 定位带判据安全假 / the safe false
    RETURN; // 早退（输出保持安全零）/ return early
END_IF

// 段 2｜防摆补偿叠加（相位对消，增益负值回拉语义，边界四）/ segment 2, the anti sway compensation
IF bAntiSwayEn THEN // 防摆使能 / the anti sway enabled
    fCorr := (fK1 * fAngDeg) + (fK2 * fAngVelDegS); // 相位对消补偿量 / the phase cancellation compensation
END_IF
_fV := fVcmd + fCorr; // 叠加 / the superposition

// 段 3｜输出钳位（±fVmax 单点回夹，边界二）/ segment 3, the outlet clamp
IF _fV > fVmax THEN // 上越界 / above the ceiling
    _fV := fVmax; // 夹到上界 / clamp to the ceiling
    bClamped := TRUE; // 信息级 / informational
ELSIF _fV < -fVmax THEN // 下越界 / below the floor
    _fV := -fVmax; // 夹到下界 / clamp to the floor
    bClamped := TRUE; // 信息级 / informational
END_IF

// 段 4｜定位带判据与统一出口（双模切换，边界三）/ segment 4, the positioning band and the outlet
bInPosBand := (ABS(fAngDeg) < fPosAngTol) AND (ABS(fAngVelDegS) < fPosVelTol); // 双容差判据 / the dual tolerance verdict
IF bEnable THEN // 输出使能 / the outlet enabled
    fVout := _fV; // 补偿速度直通 / the compensated pass through
    bValid := TRUE; // 可用 / usable
ELSE // 失能：安全侧零速显式降级（R191 降级显式声明）/ disabled, the explicit safe zero downgrade
    fVout := 0.0; // 零速 / the zero velocity
    bValid := FALSE; // 可用降假 / drop the valid
END_IF
END_FUNCTION_BLOCK

(* ---- FB_DL_CrossCorrelationDelay.st ---- *)
(*
  FB_DL_CrossCorrelationDelay  —  互相关时延估计（滑动窗 + 抛物线插值）/ Cross-correlation delay estimator
  分类 Category : DL_Algo
  码位 Code     : 16#02_3_85
  版本 Version  : 1.0.0
  来源 Source   : t2-4-s7-motion — IEC 61131-3 标准语义的道莅防御性实现
  溯源 Origin   : clean-room 实现，滑动互相关与三点抛物线亚采样插值公开语义，未复制任何源码行
                  （依赖语义对齐 FB_DL_MedianFilter / FB_DL_LowPassFilter：前端滤波由调用方承载，本件不做滤波）
  功能 Function : 1) 输入缓冲以 [0] 为最新采样点，FB 内部维护 nWindowSize 深双路滑动窗（去均值后互相关）；
                  2) 在 |lag| <= nMaxLagSamples 内取互相关峰值，三点抛物线插值得亚采样滞后 fDelayS（s，负 = 超前）；
                  3) fPeakCorr < fConfidenceMin 判不可信不出时延结论；eState: Fill/Search/Locked/Fault。
  边界 Boundary : ① fSampleDt <= 0 / nWindowSize < 16 / 2·nMaxLagSamples >= nWindowSize / 窗超数组上界 判组态错进 Fault；
                  ② 缓冲未填满时 bWindowFull := FALSE 且不出时延结论（fDelayS 维持 0）；
                  ③ 参考信号方差 < 1E-12 判「激励不足」置码且 bValid := FALSE（不输出随机滞后）；
                  ④ 峰值落窗边界（|lag| = nMaxLagSamples）判「滞后超窗」置码而非当有效值；
                  ⑤ 解除式自证：Fault 退出 = bReset 上升沿 AND 组态三参数合法（引脚均可满足，R28-1）；
                  ⑥ 未知状态由 CASE ELSE 拦截进 Fault（兜底置码）。
  依赖 Depends  : 仅 Standard.library（ABS）；前端滤波语义对齐 FB_DL_MedianFilter / FB_DL_LowPassFilter（已注册，不实例化）
  码表 Error codes（本件格 02_3_85，子码步进 +0x100）:
    16#0002_0185 信息级：参考激励不足（方差 < 1E-12），不出时延结论
    16#0002_0285 故障级：组态非法（dt <= 0 / 窗 < 16 / 2·maxLag >= 窗 / 窗超数组上界），锁存至复位
    16#0002_0385 信息级：峰值落窗边界（|lag| = maxLag），判滞后超窗
    16#0002_0485 信息级：置信度不足（fPeakCorr < fConfidenceMin），bValid = FALSE
    16#0002_0585 故障级：状态机落 ELSE 兜底（非法相位 ID）

  修订历史 Revision :
    2026-11-18  v1.0.0  R38 首版
*)

TYPE E_DL_XCorrState :
(
    eFill   := 0,   // 填窗：滑动窗未满，不出结论 / Filling, window not yet full
    eSearch := 10,  // 搜索：逐拍互相关寻峰 / Searching, per-scan peak search
    eLocked := 20,  // 锁定：峰值过置信门限，时延有效 / Locked, peak above confidence
    eFault  := 90   // 故障：组态错锁存，等复位 / Fault, latched until reset
);
END_TYPE

FUNCTION_BLOCK FB_DL_CrossCorrelationDelay
VAR_INPUT
    afSignalRef    : ARRAY[0..127] OF REAL;   // 参考信号缓冲，[0] = 本拍最新采样 / Reference buffer, index 0 is newest
    afSignalFb     : ARRAY[0..127] OF REAL;   // 反馈信号缓冲，[0] = 本拍最新采样 / Feedback buffer, index 0 is newest
    nWindowSize    : INT;                     // 相关窗长 [点]，域 16..128 / Correlation window length
    fSampleDt      : REAL;                    // 采样间隔 [s]，域 > 0 / Sample interval
    nMaxLagSamples : INT;                     // 最大滞后 [点]，域 0..63 且 2 倍 < 窗长 / Maximum lag in samples
    fConfidenceMin : REAL;                    // 置信度门限 [无量纲 0..1] / Minimum peak correlation
    bReset         : BOOL := FALSE;           // 复位（Fault 退出唯一路径）/ Reset, sole fault exit
END_VAR
VAR_OUTPUT
    fDelayS        : REAL;                    // 时延 [s]，负 = 超前 / Estimated delay, negative means lead
    fPeakCorr      : REAL;                    // 归一化峰值相关 [-1..1] / Normalized peak correlation
    bValid         : BOOL;                    // 时延结论有效 / Delay verdict valid
    bWindowFull    : BOOL;                    // 滑动窗已填满 / Window full flag
    nErrId         : UDINT;                   // 事件码，0 = 无事件 / Event code, 0 = none
    eState         : E_DL_XCorrState;         // 状态出口，段尾单点映射 / State outlet, mapped at the tail
END_VAR
VAR
    tonFaultWatch : TON;                       // 故障态驻留观察窗，自复位（段 0 无条件刷新）/ Fault dwell observer, self-resetting
    rtReset       : R_TRIG;                    // 复位上升沿 / Reset rising edge
    _eState       : E_DL_XCorrState := E_DL_XCorrState.eFill;   // 内部相位（CASE 唯一写入目标）/ Internal phase
    _arRefWin     : ARRAY[0..127] OF REAL;     // 参考滑动窗 / Reference sliding window
    _arFbWin      : ARRAY[0..127] OF REAL;     // 反馈滑动窗 / Feedback sliding window
    _arCorr       : ARRAY[0..127] OF REAL;     // 各 lag 相关系数（下标 = lag + 64）/ Correlation per lag, index = lag + 64
    _nFill        : INT;                       // 已填点数 [点] / Filled sample count
    _nPeakLag     : INT;                       // 峰值 lag [点] / Peak lag
    _nLag         : INT;                       // lag 循环计数 / Lag loop counter
    _nK           : INT;                       // 窗内循环计数 / Window loop counter
    _uFault       : UDINT;                     // 故障码锁存 / Latched fault code
    _uInfo        : UDINT;                     // 信息码，每拍重算 / Info code, recomputed per scan
    _bFault       : BOOL;                      // 故障锁存位 / Latched fault bit
    _bCfgBad      : BOOL;                      // 组态非法聚合 / Configuration invalid aggregate
    _rRefMean     : LREAL;                     // 参考窗均值 / Reference window mean
    _rFbMean      : LREAL;                     // 反馈窗均值 / Feedback window mean
    _rRefVar      : LREAL;                     // 参考窗方差 / Reference window variance
    _rFbVar       : LREAL;                     // 反馈窗方差 / Feedback window variance
    _rCross       : LREAL;                     // 交叉累加暂存 / Cross accumulation scratch
    _rPeak        : LREAL;                     // 峰值相关 / Peak correlation
    _rCm1, _rC0, _rCp1 : LREAL;                // 抛物线三点 / Parabola three points
    _rShift       : LREAL;                     // 亚采样偏移 [点] / Sub-sample shift
END_VAR
VAR CONSTANT
    nWinMin  : INT   := 16;       // 最小窗长 [点] / Minimum window length
    nWinMax  : INT   := 128;      // 数组上界 [点] / Array upper bound
    nLagBase : INT   := 64;       // lag 下标基准（数组下标 = lag + 64）/ Lag index base
    rVarFloor: LREAL := 1.0E-12;  // 激励方差下限 / Excitation variance floor
    rWatchPt : TIME  := T#2S;     // 故障观察窗 [ms]，自复位节拍 / Fault watch window, self-resetting
END_VAR

(* —— 段 0：定时器与边沿无条件周期刷新（R182：调用语句不得置于 IF/CASE 内） —— *)
rtReset(CLK := bReset);                                     // 复位上升沿，每拍必调
tonFaultWatch(IN := (NOT tonFaultWatch.Q), PT := rWatchPt); // 观察窗自复位节拍（表达式入参，非 IF 内）

(* —— 段 1：单拍量预清零（锁存量 _uFault/_bFault/_nFill/_arWin 不入清单，R187①） —— *)
_uInfo    := 16#0000_0000;     // 信息码每拍重算
bValid    := FALSE;            // 结论缺省无效
nErrId    := 16#0000_0000;     // 事件码缺省无事件

(* —— 段 2：组态域闸（覆盖全部参与判据换算的引脚，R151） —— *)
_bCfgBad := FALSE;             // 组态非法预清零（每拍重算，Fault 锁存不受影响）
IF LREAL(fSampleDt) <= 0.0 THEN
    _bCfgBad := TRUE;          // 采样间隔非法
END_IF
IF (nWindowSize < nWinMin) OR (nWindowSize > nWinMax) THEN
    _bCfgBad := TRUE;          // 窗长越域
END_IF
IF (nMaxLagSamples < 0) OR ((2 * nMaxLagSamples) >= nWindowSize) THEN
    _bCfgBad := TRUE;          // 滞后窗不得吃掉相关样本（规格强制）
END_IF
IF _bCfgBad THEN
    _uFault  := 16#0002_0285;  // 故障级：组态非法
    _bFault  := TRUE;          // 锁存（解除式自证：bReset AND 组态合法）
    _eState  := E_DL_XCorrState.eFault;
END_IF

(* —— 段 3：复位沿（Fault 解除唯一路径：bReset AND 组态合法） —— *)
IF rtReset.Q THEN
    IF (NOT _bCfgBad) THEN
        _bFault  := FALSE;                 // 清故障锁存位
        _uFault  := 16#0000_0000;          // 清锁存码
        _eState  := E_DL_XCorrState.eFill; // 回填窗相重新开始
        _nFill   := 0;                     // 填充计数清零
        fDelayS  := 0.0;                   // 时延结论清零
        fPeakCorr := 0.0;                  // 峰值清零
    END_IF
END_IF

(* —— 段 4：滑动窗移位入队（每拍执行，Fault 相冻结不采集） —— *)
IF _eState <> E_DL_XCorrState.eFault THEN
    FOR _nK := (nWinMax - 1) TO 1 BY -1 DO
        _arRefWin[_nK] := _arRefWin[_nK - 1];   // 参考窗右移
        _arFbWin[_nK]  := _arFbWin[_nK - 1];    // 反馈窗右移
    END_FOR
    _arRefWin[0] := afSignalRef[0];             // 最新采样入队（[0] = 本拍最新）
    _arFbWin[0]  := afSignalFb[0];
    IF _nFill < nWinMax THEN
        _nFill := _nFill + 1;                   // 填充计数（上限守卫，不回绕）
    END_IF
END_IF
bWindowFull := _nFill >= nWindowSize;           // 窗满标志（窗长已闸 <= 128）

(* —— 段 5：相位机（只做迁移与计算；出口在段 8） —— *)
CASE _eState OF

E_DL_XCorrState.eFill:
    IF bWindowFull THEN
        _eState := E_DL_XCorrState.eSearch;     // 窗满：进搜索相
    END_IF

E_DL_XCorrState.eSearch:
    IF NOT bWindowFull THEN
        _eState := E_DL_XCorrState.eFill;       // 组态变更窗长变大：回填窗相
    ELSE
        (* —— 去均值与方差（分母 nWindowSize 已闸 >= 16） —— *)
        _rRefMean := 0.0;  _rFbMean := 0.0;
        FOR _nK := 0 TO (nWindowSize - 1) DO
            _rRefMean := _rRefMean + LREAL(_arRefWin[_nK]);
            _rFbMean  := _rFbMean  + LREAL(_arFbWin[_nK]);
        END_FOR
        _rRefMean := _rRefMean / LREAL(nWindowSize);
        _rFbMean  := _rFbMean  / LREAL(nWindowSize);
        _rRefVar  := 0.0;  _rFbVar := 0.0;
        FOR _nK := 0 TO (nWindowSize - 1) DO
            _rRefVar := _rRefVar + (LREAL(_arRefWin[_nK]) - _rRefMean) * (LREAL(_arRefWin[_nK]) - _rRefMean);
            _rFbVar  := _rFbVar  + (LREAL(_arFbWin[_nK])  - _rFbMean)  * (LREAL(_arFbWin[_nK])  - _rFbMean);
        END_FOR
        _rRefVar := _rRefVar / LREAL(nWindowSize);
        _rFbVar  := _rFbVar  / LREAL(nWindowSize);
        IF _rRefVar < rVarFloor THEN
            _uInfo := 16#0002_0185;             // 信息级：参考激励不足
            fPeakCorr := 0.0;                   // 不输出随机滞后
        ELSE
            (* —— 滑动互相关（lag ∈ [−maxLag, +maxLag]，重叠区去均值归一化） —— *)
            _rPeak := -2.0;                     // 峰值暂存（相关系数域 [-1,1]，取超域初值）
            _nPeakLag := 0;
            FOR _nLag := -nMaxLagSamples TO nMaxLagSamples DO
                _rCross := 0.0;
                FOR _nK := 0 TO (nWindowSize - 1 - ABS(_nLag)) DO
                    _rCross := _rCross
                        + (LREAL(_arRefWin[_nK]) - _rRefMean)
                        * (LREAL(_arFbWin[_nK + _nLag]) - _rFbMean);   // 参考滞后 _nLag 拍的交叉积
                END_FOR
                _arCorr[_nLag + nLagBase] := REAL(_rCross
                    / MAX(SQRT(_rRefVar * _rFbVar) * LREAL(nWindowSize - ABS(_nLag)), rVarFloor));  // 归一化（分母已闸）
                IF LREAL(_arCorr[_nLag + nLagBase]) > _rPeak THEN
                    _rPeak := LREAL(_arCorr[_nLag + nLagBase]);        // 峰值刷新
                    _nPeakLag := _nLag;                                 // 峰值 lag 记录
                END_IF
            END_FOR
            fPeakCorr := REAL(_rPeak);
            (* —— 边界峰值 = 滞后超窗：判码不出有效值（规格强制） —— *)
            IF ABS(_nPeakLag) >= nMaxLagSamples THEN
                _uInfo := 16#0002_0385;         // 信息级：峰值落窗边界
            ELSIF _rPeak < LREAL(fConfidenceMin) THEN
                _uInfo := 16#0002_0485;         // 信息级：置信度不足
            ELSE
                (* —— 三点抛物线亚采样插值（峰值在开区间内，三点必在 lag 表内） —— *)
                _rCm1 := LREAL(_arCorr[_nPeakLag - 1 + nLagBase]);   // lag−1 相关系数
                _rC0  := LREAL(_arCorr[_nPeakLag     + nLagBase]);   // lag   相关系数
                _rCp1 := LREAL(_arCorr[_nPeakLag + 1 + nLagBase]);   // lag+1 相关系数
                IF ABS(_rCm1 - 2.0 * _rC0 + _rCp1) > rVarFloor THEN
                    _rShift := 0.5 * (_rCm1 - _rCp1) / (_rCm1 - 2.0 * _rC0 + _rCp1);   // 抛物线顶点偏移（分母已闸）
                ELSE
                    _rShift := 0.0;             // 三点共线：退化为整数 lag
                END_IF
                fDelayS := REAL((LREAL(_nPeakLag) + _rShift) * LREAL(fSampleDt));   // 亚采样时延 [s]
                bValid  := TRUE;                // 结论有效
                _eState := E_DL_XCorrState.eLocked;   // 过门限：进锁定相
            END_IF
        END_IF
    END_IF

E_DL_XCorrState.eLocked:
    IF NOT bWindowFull THEN
        _eState := E_DL_XCorrState.eFill;       // 组态变更：回填窗相
        bValid  := FALSE;                       // 锁定值作废
    ELSE
        (* —— 锁定相维持结论并继续逐拍复算（复算逻辑与搜索相同，保持时延新鲜度） —— *)
        _rRefMean := 0.0;  _rFbMean := 0.0;
        FOR _nK := 0 TO (nWindowSize - 1) DO
            _rRefMean := _rRefMean + LREAL(_arRefWin[_nK]);
            _rFbMean  := _rFbMean  + LREAL(_arFbWin[_nK]);
        END_FOR
        _rRefMean := _rRefMean / LREAL(nWindowSize);
        _rFbMean  := _rFbMean  / LREAL(nWindowSize);
        _rRefVar  := 0.0;  _rFbVar := 0.0;
        FOR _nK := 0 TO (nWindowSize - 1) DO
            _rRefVar := _rRefVar + (LREAL(_arRefWin[_nK]) - _rRefMean) * (LREAL(_arRefWin[_nK]) - _rRefMean);
            _rFbVar  := _rFbVar  + (LREAL(_arFbWin[_nK])  - _rFbMean)  * (LREAL(_arFbWin[_nK])  - _rFbMean);
        END_FOR
        _rRefVar := _rRefVar / LREAL(nWindowSize);
        _rFbVar  := _rFbVar  / LREAL(nWindowSize);
        IF _rRefVar < rVarFloor THEN
            _uInfo := 16#0002_0185;             // 信息级：激励不足（锁定值维持，bValid 置 FALSE）
            bValid := FALSE;
        ELSE
            _rPeak := -2.0;
            _nPeakLag := 0;
            FOR _nLag := -nMaxLagSamples TO nMaxLagSamples DO
                _rCross := 0.0;
                FOR _nK := 0 TO (nWindowSize - 1 - ABS(_nLag)) DO
                    _rCross := _rCross
                        + (LREAL(_arRefWin[_nK]) - _rRefMean)
                        * (LREAL(_arFbWin[_nK + _nLag]) - _rFbMean);
                END_FOR
                _arCorr[_nLag + nLagBase] := REAL(_rCross
                    / MAX(SQRT(_rRefVar * _rFbVar) * LREAL(nWindowSize - ABS(_nLag)), rVarFloor));
                IF LREAL(_arCorr[_nLag + nLagBase]) > _rPeak THEN
                    _rPeak := LREAL(_arCorr[_nLag + nLagBase]);
                    _nPeakLag := _nLag;
                END_IF
            END_FOR
            fPeakCorr := REAL(_rPeak);
            IF ABS(_nPeakLag) >= nMaxLagSamples THEN
                _uInfo := 16#0002_0385;         // 信息级：滞后超窗（锁定值维持，bValid 置 FALSE）
                bValid := FALSE;
            ELSIF _rPeak < LREAL(fConfidenceMin) THEN
                _uInfo := 16#0002_0485;         // 信息级：置信度不足
                bValid := FALSE;
            ELSE
                _rCm1 := LREAL(_arCorr[_nPeakLag - 1 + nLagBase]);
                _rC0  := LREAL(_arCorr[_nPeakLag     + nLagBase]);
                _rCp1 := LREAL(_arCorr[_nPeakLag + 1 + nLagBase]);
                IF ABS(_rCm1 - 2.0 * _rC0 + _rCp1) > rVarFloor THEN
                    _rShift := 0.5 * (_rCm1 - _rCp1) / (_rCm1 - 2.0 * _rC0 + _rCp1);
                ELSE
                    _rShift := 0.0;
                END_IF
                fDelayS := REAL((LREAL(_nPeakLag) + _rShift) * LREAL(fSampleDt));   // 时延逐拍刷新
                bValid  := TRUE;                // 结论维持有效
            END_IF
        END_IF
    END_IF

E_DL_XCorrState.eFault:
    ;                                           // 故障相：等复位沿（段 3 承载解除，无动作）

ELSE
    _uFault := 16#0002_0585;                    // 故障级：非法相位 ID 兜底
    _bFault := TRUE;                            // 锁存
    _eState := E_DL_XCorrState.eFault;          // 强制回故障相

END_CASE

(* —— 段 6：出口单点映射（名实同源；锁存码回放，禁同拍抹除） —— *)
eState := _eState;                              // 状态出口单点映射
IF _bFault THEN
    nErrId := _uFault;                          // 故障锁存码回放（不在故障相按当下输入重推）
    bValid := FALSE;                            // 故障相结论无效（安全侧）
ELSE
    nErrId := _uInfo;                           // 信息码
END_IF

END_FUNCTION_BLOCK

(* ---- FB_DL_CusumMonitor.st ---- *)
(*==============================================================================
 * 组件名称 (Component)  : FB_DL_CusumMonitor
 * 所属子库 (Sublibrary) : DL_Algo
 * 当前版本 (Version)    : 1.0.0
 * 兼容性   (Platform)   : CODESYS 3.5+ / TwinCAT 3 / 汇川 InoProShop / 施耐德 Machine Expert
 *                         仅依赖 Standard.library（ABS / MAX），零厂商私有库
 * 功能描述 (Function)   : 双侧 CUSUM 累积和监视（Page 型决策区间）：
 *                           fCpos = MAX(0, fCpos + (fSample − fTarget − fK))
 *                           fCneg = MAX(0, fCneg + (fTarget − fSample − fK))
 *                         正/负决策区间下限钳零（防负累加，规格指定）；累计和
 *                         达决策限 fH（>= 容差判）置 bPosAlarm / bNegAlarm
 *                         （电平输出，回落自动撤销，不锁存）；bReset 上升沿清
 *                         双累计与计数。非有限样本跳过递推并计数置信息码
 *                         eSampleSkip（规格指定）。
 * 接口     (Interface)  : 输入 fSample 观测样本、fTarget 目标均值、fK 容许限
 *                         （域 > 0）、fH 决策限（域 > 0）、bReset 复位；
 *                         输出 fCpos 正向累计和、fCneg 负向累计和、bPosAlarm
 *                         正偏报警（电平）、bNegAlarm 负偏报警（电平）、
 *                         uSkipCnt 非有限样本跳过计数、eErrCode 错误码、
 *                         bError 故障标志。
 * 边界     (Boundary)   : ① **属主边界（写死）：本件只做 CUSUM 递推与双侧判限，
 *                         不接管报警管理、不归一化样本**；报警归集归
 *                         `FB_DL_AlarmManager`。
 *                         ② 递推钳零：MAX(0, ·) 使区间单调不下降且非负，
 *                         结构性防负累加（规格指定口径）。
 *                         ③ 报警判据 fCpos >= fH 用容差比较（禁浮点 =），
 *                         电平语义（回落撤销）写入头注释，非锁存。
 *                         ④ 非有限样本（R79 双判）跳过递推：双累计不被污染，
 *                         uSkipCnt 防回绕递增，信息码不置 bError。
 *                         ⑤ 组态闸：fK <= 0 或 fH <= 0 → 锁存故障，双累计
 *                         冻结、报警出口安全侧 FALSE，解除沿 = bReset 上升沿
 *                         （故障级码配对 bError，R45）。
 *                         ⑥ 零全局耦合（无 GVL / VAR_EXTERNAL / 物理地址）。
 * 分工声明 (Scope)      : 与 `FB_DL_Integrator` 分工：无界积分归那件、钳零双侧
 *                         决策区间归本件；与 `FB_DL_EtchEndpointTrend` 分工：
 *                         工艺终点趋势归那件。
 * 来源标签 (Source Tag) : 自研线（Page CUSUM 为公开统计过程控制定义 clean-room）
 * 码表     (Codes)      : 本件不占用任何全局数字码位。出口为 LREAL 累计组 +
 *                         BOOL 报警组 + UDINT 计数 + ENUM 错误码；数字码位待
 *                         主控收口阶段统一派号。
 * 红线自检 (Redline)    : R1 ✓ 零 GVL/VAR_EXTERNAL ｜ R2 ✓ 零 %I/%Q/%M ｜ R3 ✓ 纯 IEC 61131-3
 *                         R4 ✓ 钳零递推 + 非有限跳过 + 组态锁存 ｜ R5 ✓ 声明逐行同行双语注释
 *                         R6 N/A（无 ENUM 状态机） ｜ R7 ✓ 一 R_TRIG 段 0 无条件刷新
 * 修订历史 (Revision)   : 2026-11-20  v1.0.0  R50 首版（批次 2 · 序号 6）
 * 验收向量 (Acceptance) : ① fTarget=10, fK=0.5, fH=5，样本 12,12,12,12 →
 *                         fCpos = 1.5, 3.0, 4.5, 6.0，第 4 拍 6.0 >= 5 →
 *                         bPosAlarm=TRUE，fCneg 恒 0；② 样本 8,8 → fCneg =
 *                         2.5, 5.0，第 2 拍 bNegAlarm=TRUE，fCpos 恒 0；
 *                         ③ fK=0 → 锁存故障 eCfgBad，出口冻结；
 *                         ④ 样本 NaN → uSkipCnt+1，eErrCode=eSampleSkip，
 *                         累计不变。
 *==============================================================================*)

(*-----------------------------------------------------------------------------
 * 枚举: E_DL_CusumErr（错误码；信息级不置 bError，故障级恒伴 bError=TRUE）
 *----------------------------------------------------------------------------*)
TYPE E_DL_CusumErr :
(
    eOk         := 0,   // 正常 / Normal
    eCfgBad     := 1,   // 故障级：组态非法（fK/fH 域） / Fault: illegal configuration
    eSampleSkip := 2    // 信息级：非有限样本跳过（见 uSkipCnt） / Info: non-finite sample skipped
);
END_TYPE

FUNCTION_BLOCK FB_DL_CusumMonitor
VAR_INPUT
    fSample : LREAL := 0.0;           // 观测样本 [工程单位] / Observed sample
    fTarget : LREAL := 0.0;           // 目标均值（与样本同工程单位） / Target mean, same engineering unit
    fK      : LREAL := 0.5;           // 容许限（偏移容忍），域 > 0 [工程单位] / Allowance, must be > 0
    fH      : LREAL := 5.0;           // 决策限（累计和阈值），域 > 0 [工程单位] / Decision limit, must be > 0
    bReset  : BOOL := FALSE;          // 复位，上升沿清双累计与跳过计数 [-] / Reset, rising edge clears accumulators
END_VAR
VAR_OUTPUT
    fCpos     : LREAL;                // 正向累计和（下限钳零） [工程单位] / Positive cumulative sum, floored at zero
    fCneg     : LREAL;                // 负向累计和（下限钳零） [工程单位] / Negative cumulative sum, floored at zero
    bPosAlarm : BOOL;                 // 正偏报警电平（fCpos >= fH） [-] / Positive alarm level
    bNegAlarm : BOOL;                 // 负偏报警电平（fCneg >= fH） [-] / Negative alarm level
    uSkipCnt  : UDINT := 0;           // 非有限样本跳过计数（防回绕） [个] / Skipped-sample counter
    eErrCode  : E_DL_CusumErr;        // 错误码出口 / Error code outlet
    bError    : BOOL;                 // 故障标志（组态锁存） [-] / Error flag, latched
END_VAR
VAR
    _fCpos    : LREAL := 0.0;         // 正向累计锁存（冻结源，与出口同源） / Positive sum latch
    _fCneg    : LREAL := 0.0;         // 负向累计锁存 / Negative sum latch
    _bNonFin  : BOOL;                 // 样本非有限当拍量 [-] / Sample non-finite this scan
    _bCfgBad  : BOOL;                 // 组态非法当拍量 [-] / Illegal configuration this scan
    _bErrLatch: BOOL;                 // 组态故障锁存位（解除沿 = bReset 上升沿） / Latched config fault
    rtReset   : R_TRIG;               // 复位沿实例，段 0 无条件调用 / Reset edge instance
END_VAR
VAR CONSTANT
    DL_CSM_ZERO : LREAL := 0.0;       // 钳零下限与判零基准 [工程单位] / Zero floor and non-finite base
    DL_CSM_UDMAX: UDINT := 4294967295;   // 跳过计数饱和点（防回绕） [个] / Skip counter saturation ceiling
END_VAR

(* —— 段 0：非有限判 + 组态闸 + 沿刷新 —— *)
_bNonFin := (fSample <> fSample) OR ((fSample - fSample) <> DL_CSM_ZERO);   // 样本非有限（R79 双判） / Sample non-finite
_bCfgBad := (fK <= DL_CSM_ZERO) OR (fH <= DL_CSM_ZERO);                     // 组态域闸（fK/fH 须正） / Configuration gate
rtReset(CLK := bReset);                            // 复位沿，每拍必调 / Reset edge, every scan

(* —— 段 1：复位沿（清双累计与跳过计数；先于故障锁存判定，复位语义优先） —— *)
IF rtReset.Q THEN
    _fCpos := DL_CSM_ZERO;                         // 清正向累计（规格：复位沿清双累计） / Clear positive sum
    _fCneg := DL_CSM_ZERO;                         // 清负向累计 / Clear negative sum
    uSkipCnt := 0;                                 // 清跳过计数 / Clear skip counter
    _bErrLatch := FALSE;                           // 清组态锁存（R188 声明：解除沿 = bReset 上升沿） / Clear cfg latch
END_IF
IF _bCfgBad AND (NOT _bErrLatch) THEN
    _bErrLatch := TRUE;                            // 锁存 / Latch
END_IF

(* —— 段 2：CUSUM 递推（组态故障期冻结；非有限样本跳过） —— *)
IF (NOT _bErrLatch) AND (NOT _bNonFin) THEN
    _fCpos := MAX(DL_CSM_ZERO, _fCpos + (fSample - fTarget - fK));   // 正向递推钳零 / Positive recursion floored
    _fCneg := MAX(DL_CSM_ZERO, _fCneg + (fTarget - fSample - fK));   // 负向递推钳零 / Negative recursion floored
ELSIF (NOT _bErrLatch) AND _bNonFin THEN
    IF uSkipCnt < DL_CSM_UDMAX THEN
        uSkipCnt := uSkipCnt + 1;                  // 跳过计数防回绕递增 / Skip counter increment
    END_IF
END_IF

(* —— 段 3：出口单点映射（名实双出口同源，R191） —— *)
fCpos := _fCpos;                                   // 正向累计出口 / Positive sum outlet
fCneg := _fCneg;                                   // 负向累计出口 / Negative sum outlet
IF _bErrLatch THEN
    bPosAlarm := FALSE;                            // 故障安全侧：报警出口 FALSE / Fault safe side
    bNegAlarm := FALSE;                            // 故障安全侧：负偏报警出口 FALSE / Fault safe side for negative alarm
    bError := TRUE;                                // 故障标志（R45 配对） / Error flag
    eErrCode := E_DL_CusumErr.eCfgBad;             // 故障级码 / Fault code
ELSE
    bPosAlarm := _fCpos >= fH;                     // 报警电平（容差域 >= 判，禁 =） / Positive alarm level
    bNegAlarm := _fCneg >= fH;                     // 负偏报警电平 / Negative alarm level
    IF _bNonFin THEN
        eErrCode := E_DL_CusumErr.eSampleSkip;     // 信息级（不置 bError） / Info code
    ELSE
        eErrCode := E_DL_CusumErr.eOk;             // 正常 / Normal
    END_IF
    bError := FALSE;                               // 无故障级条件 / No fault
END_IF

END_FUNCTION_BLOCK

(* ---- FB_DL_DeadbandFilter.st ---- *)
(*==============================================================================
 * 组件名称 (Component)  : FB_DL_DeadbandFilter
 * 所属子库 (Sublibrary) : DL_Algo
 * 当前版本 (Version)    : 1.0.0
 * 兼容性   (Platform)   : CODESYS 3.5+ / TwinCAT 3 / 汇川 InoProShop / 施耐德 Machine Expert
 *                         仅依赖 Standard.library（ABS），零厂商私有库
 * 功能描述 (Function)   : **双向死区 + 输出保持**（有状态件）。规则：
 *                           |fIn - fOut| > fDeadband → fOut := fIn（采纳），bUpdated=TRUE；
 *                           否则 fOut 保持不动（抑制抖振），bUpdated=FALSE。
 *                         与无状态单值死区 FC（FC_DL_Deadband）的差别：那件每拍独立判断
 *                         「输入是否落在死区内并输出 0 或原值」，**不记忆历史**；
 *                         本件记忆上一输出，死区判定以**上一输出**为基准，
 *                         故能彻底消除阈值附近的来回抖动（迟滞特性），
 *                         但代价是引入 ≤ fDeadband 的稳态静差（现场需知悉）。
 * 接口     (Interface)  : 输入 bEnable 使能、bReset 复位输出到当前输入、fIn 采样输入 [EU]、
 *                         fDeadband 双向死区宽度 [EU]（>= 0）；
 *                         输出 fOut 输出值（保持语义） [EU]、bUpdated 本拍是否更新、
 *                         fDeviation 当前偏差 |fIn-fOut| [EU]、bValid 输出有效、
 *                         bError 故障标志、uErrorId 故障码。
 * 边界     (Boundary)   : ① 属主边界：只做死区保持，不做平滑 / 限速 / 量化（另件）。
 *                         ② fDeadband < 0 → 故障级 16#0008_0003（负死区会放大抖振，禁止钳位后静默放行）。
 *                         ③ fDeadband = 0 → 退化为直通（任何偏差都采纳），合法。
 *                         ④ 非有限防御：fIn 与 fDeadband 逐一枚举，命中即故障态 16#0008_0002，
 *                         输出冻结（不推 0）。
 *                         ⑤ 恢复路径：bEnable=FALSE 或 bReset=TRUE 均可解除故障态。
 *                         ⑥ 零全局耦合（无 GVL / VAR_EXTERNAL / 物理地址）。
 * 分工声明 (Scope)      : 与无状态 `FC_DL_Deadband` 分工：单值死区归那件、带记忆的
 *                         死区保持归本件；与 `FB_DL_QuantizeFilter` 分工：量化+回差归那件。
 * 来源标签 (Source Tag) : 原创实现（无外部代码引入）
 * 码表     (Codes)      : 16#0008_0000 无故障 / 16#0008_0002 入参非有限（故障级）/
 *                         16#0008_0003 死区为负（故障级）/ 16#0008_0005 非法状态（故障级）。
 * 红线自检 (Redline)    : R1 ✓ 零 GVL/VAR_EXTERNAL ｜ R2 ✓ 零 %I/%Q/%M ｜ R3 ✓ 纯 IEC 61131-3
 *                         R4 ✓ 双浮点入参非有限判 + 死区符号域闸 + 无除法 ｜ R5 ✓ 声明逐行同行双语注释
 *                         R6 ✓ 四态 ENUM + CASE + ELSE 兜底 ｜ R7 N/A（无 TON / 边沿实例）
 * 修订历史 (Revision)   : 2026-11-23  v1.0.0  R77 首版（批次 B3 · 序号 14）
 * 验收向量 (Acceptance) : ① fDeadband=2.0，fIn=10.0（fOut 初 0）→ |10-0|=10 > 2 → fOut=10.0, bUpdated=TRUE；
 *                         ② 随后 fIn=11.0 → |11-10|=1 <= 2 → fOut 保持 10.0, bUpdated=FALSE；
 *                         ③ 随后 fIn=12.5 → |12.5-10|=2.5 > 2 → fOut=12.5, bUpdated=TRUE；
 *                         ④ fDeadband=0.0 → 任何变化都采纳（直通），fOut=fIn；
 *                         ⑤ fDeadband=-1.0 → uErrorId=16#0008_0003，bError=TRUE，fOut 冻结。
 *==============================================================================*)

(*-----------------------------------------------------------------------------
 * 枚举: E_DL_DeadbandState（死区保持状态机，归属 DL_Algo，与本件同文件，全库唯一属主）
 *----------------------------------------------------------------------------*)
TYPE E_DL_DeadbandState :
(
    eInit  := 0,    // 首扫 / 复位后：输出直取输入 / First scan or after reset: output follows input
    eRun   := 10,   // 运行态：死区外采纳、死区内保持 / Running: adopt outside band, hold inside band
    eHoldF := 20,   // 保持态：未使能，输出冻结 / Hold: disabled, output frozen
    eFault := 99    // 故障态：输出冻结，等待 bEnable 跌落或 bReset / Fault: frozen until cleared
);
END_TYPE

FUNCTION_BLOCK FB_DL_DeadbandFilter
VAR_INPUT
    bEnable   : BOOL := FALSE;   // 使能，FALSE 冻结输出 / Enable, FALSE freezes output
    bReset    : BOOL := FALSE;   // 复位输出到当前输入（单拍有效） / Reset output to current input, single scan
    fIn       : LREAL := 0.0;    // 采样输入 [EU] / Sampling input [EU]
    fDeadband : LREAL := 0.5;    // 双向死区宽度，必须 >= 0 [EU] / Two-sided deadband width, must be non-negative [EU]
END_VAR
VAR_OUTPUT
    fOut      : LREAL;   // 输出值（死区内保持） [EU] / Output value, held inside the deadband [EU]
    bUpdated  : BOOL;    // 本拍是否更新输出 [-] / Whether the output updated this scan
    fDeviation: LREAL;   // 当前偏差 |fIn - fOut| [EU] / Current deviation [EU]
    bValid    : BOOL;    // 输出有效标志 [-] / Output valid flag
    bError    : BOOL;    // 故障标志，与 uErrorId 联动 [-] / Fault flag coupled with uErrorId
    uErrorId  : UDINT;   // 故障码，0 = 无故障 [-] / Error code, zero means healthy
END_VAR
VAR
    _bNonFin : BOOL;               // 入参非有限标志 [-] / Non-finite input flag
    eState   : E_DL_DeadbandState; // 状态机当前状态 [-] / Current state
END_VAR
VAR CONSTANT
    DL_DBF_ZERO : LREAL := 0.0;    // 零基准（含非有限判零） [-] / Zero base including non-finite probe
END_VAR

(* —— 段 1：非有限防御（fIn 与 fDeadband 逐一枚举） —— *)
uErrorId := 16#0008_0000;                          // 预置无故障 / Preset healthy
_bNonFin := (fIn <> fIn) OR ((fIn - fIn) <> DL_DBF_ZERO);              // 输入非有限 / Input non-finite
_bNonFin := _bNonFin OR (fDeadband <> fDeadband) OR ((fDeadband - fDeadband) <> DL_DBF_ZERO);  // 死区非有限
IF _bNonFin THEN
    eState   := eFault;                            // 强制故障态 / Force fault state
    uErrorId := 16#0008_0002;                      // 故障级：入参非有限 / Fault: non-finite input
END_IF

(* —— 段 2：死区符号域闸（负死区会放大抖振，必须拒绝而非钳位） —— *)
IF fDeadband < DL_DBF_ZERO THEN
    eState   := eFault;
    uErrorId := 16#0008_0003;                      // 故障级：死区为负 / Fault: negative deadband
END_IF

(* —— 段 3：复位请求 → 回首扫 —— *)
IF bReset THEN
    eState := eInit;
END_IF

(* —— 段 4：状态派生 —— *)
IF NOT bEnable THEN
    eState := eHoldF;                              // 未使能：冻结 / Disabled: freeze
ELSIF eState = eFault THEN
    eState := eFault;                              // 故障态保持 / Fault holds
ELSIF eState = eInit THEN
    eState := eInit;                               // 首扫保持一拍 / Init holds one scan
ELSE
    eState := eRun;
END_IF

(* —— 段 5：主状态机（CASE 覆盖 + ELSE 兜底） —— *)
CASE eState OF

    eInit:
        fOut       := fIn;                         // 首拍直取输入 / First scan follows input
        fDeviation := DL_DBF_ZERO;
        bUpdated   := TRUE;
        bValid     := TRUE;
        eState     := eRun;

    eRun:
        fDeviation := ABS(fIn - fOut);             // 偏差以「上一输出」为基准（迟滞核心） / Deviation versus previous output
        IF fDeviation > fDeadband THEN
            fOut     := fIn;                       // 跳出死区：采纳新值 / Outside band: adopt
            bUpdated := TRUE;
        ELSE
            (* 死区内：fOut 保持不动，不做任何改写 / Inside band: hold unchanged *)
            bUpdated := FALSE;
        END_IF
        bValid := TRUE;

    eHoldF:
        (* 未使能：输出与偏差保持上拍值 / Disabled: output and deviation frozen *)
        bUpdated := FALSE;
        bValid   := FALSE;

    eFault:
        (* 故障态：输出冻结保持上拍值（不推 0，避免下游误判为真实零） / Fault: output frozen *)
        bUpdated := FALSE;
        bValid   := FALSE;

    ELSE
        eState   := eFault;
        bUpdated := FALSE;
        bValid   := FALSE;
        uErrorId := 16#0008_0005;                  // 故障级：非法状态 / Fault: illegal state

END_CASE;

(* —— 段 6：出口映射（bError 与 uErrorId 同源；本件无信息级码） —— *)
bError := (uErrorId <> 16#0008_0000);

END_FUNCTION_BLOCK

(* ---- FB_DL_Decouple2x2.st ---- *)
(*==============================================================================
 * 组件名称 (Component)  : FB_DL_Decouple2x2
 * 所属子库 (Sublibrary) : DL_Algo
 * 当前版本 (Version)    : 1.0.0
 * 兼容性   (Platform)   : CODESYS 3.5+ / TwinCAT 3 / 汇川 InoProShop / 施耐德 Machine Expert
 *                         仅依赖 Standard.library（ABS），零厂商私有库
 * 功能描述 (Function)   : 2×2 强耦合回路静态解耦网：静态解耦注入式
 *                           fU1Eff = fU1 + fD21×fU2
 *                           fU2Eff = fU2 + fD12×fU1
 *                         fD12 / fD21 = 组态解耦系数 = Δu_i 对 j 回路的静态影响比（无量纲）。
 *                         Bristol 相对增益整定参考（写入注释供现场整定者）：
 *                           fD12 ≈ -K12/K11，fD21 ≈ -K21/K22（Kij 为开环静态增益阵元，
 *                           T21 = K12×K21/(K11×K22) 作耦合强弱组态参考，本件不计算 T 值）。
 * 接口     (Interface)  : 输入 fU1/fU2 两主控输出（0~100%）、fD12/fD21 解耦系数（无量纲，
 *                         域 |fD|<=1）、bEnable 使能、bReset 复位；输出 fU1Eff/fU2Eff
 *                         解耦后等效输出（0~100%）、bEnabled 生效指示、bCfgBad 组态非法
 *                         （锁存）、bError 故障标志。
 * 边界     (Boundary)   : ① **属主边界（写死）：本件只做静态解耦注入与输出钳位，不做动态
 *                         补偿、不接管主控 PID**；主控输出由上层 PID 件给出。
 *                         ② bEnable=FALSE 直通：fU1Eff:=fU1、fU2Eff:=fU2（不冻结历史值，
 *                         直通即语义，头注释声明）。
 *                         ③ 输出钳 [0,100%]（解耦注入可能越出主控行程，钳位防执行器饱和
 *                         反卷积）；钳位不置故障（饱和不等于故障）。
 *                         ④ 非有限输入直通拒改（fU/fD 任一非有限当拍按直通处理，R245）；
 *                         fD 非有限属组态病 → 锁存 bCfgBad。
 *                         ⑤ 解耦系数域闸：|fD12|>1 或 |fD21|>1 → 锁存 bCfgBad（反向主导
 *                         说明组态颠倒，比静默错注入危险），直通运行，解除沿 = bReset 上升沿。
 *                         ⑥ 零全局耦合（无 GVL / 无 VAR_EXTERNAL / 无物理地址）。
 * 分工声明 (Scope)      : 与 `FB_DL_CascadePid` 分工：解耦网（并联注入）≠ 串级（主从串联）；
 *                         二者可组合不可互替。
 * 来源标签 (Source Tag) : T2-1 ◐（公开 Bristol RGA 公式只借整定口径，解耦网实现自研）
 * 码表     (Codes)      : 本件不占用任何全局数字码位。出口为 LREAL 组 + BOOL 组；
 *                         数字码位待主控收口阶段统一派号。
 * 红线自检 (Redline)    : R1 ✓ 零 GVL/VAR_EXTERNAL ｜ R2 ✓ 零 %I/%Q/%M ｜ R3 ✓ 纯 IEC 61131-3
 *                         R4 ✓ 系数域闸 + 非有限直通 + 输出钳位 ｜ R5 ✓ 声明逐行同行双语注释
 *                         R6 N/A（无 ENUM 状态机） ｜ R7 ✓ 一 R_TRIG 段 0 无条件刷新
 * 修订历史 (Revision)   : 2026-11-20  v1.0.0  R48 首版（批次 2 · 序号 9）
 *                         验收向量：fD=0 → 直通；fD21=0.5、fU2=100 → U1Eff 钳 100；
 *                         |fD|=1.2 → bCfgBad 锁存直通。
 *==============================================================================*)

FUNCTION_BLOCK FB_DL_Decouple2x2
VAR_INPUT
    fU1    : LREAL := 0.0;    // 主控 1 输出（解耦前） [%] / Controller 1 output before decoupling [%]
    fU2    : LREAL := 0.0;    // 主控 2 输出（解耦前） [%] / Controller 2 output before decoupling [%]
    fD12   : LREAL := 0.0;    // 解耦系数：u1 对回路 2 的静态影响比（域 |fD|<=1） [无量纲] / Decoupling factor u1 onto loop 2
    fD21   : LREAL := 0.0;    // 解耦系数：u2 对回路 1 的静态影响比（域 |fD|<=1） [无量纲] / Decoupling factor u2 onto loop 1
    bEnable: BOOL := FALSE;   // 使能（FALSE=直通） [-] / Enable, FALSE bypasses
    bReset : BOOL := FALSE;   // 复位，上升沿清 bCfgBad 锁存 [-] / Reset, rising edge clears cfg latch
END_VAR
VAR_OUTPUT
    fU1Eff  : LREAL;          // 解耦后回路 1 等效输出（已钳 0~100%） [%] / Loop 1 effective output, clamped 0..100%
    fU2Eff  : LREAL;          // 解耦后回路 2 等效输出（已钳 0~100%） [%] / Loop 2 effective output, clamped 0..100%
    bEnabled: BOOL;           // 解耦生效指示（使能 ∧ 组态合法） [-] / Decoupling active indicator
    bCfgBad : BOOL;           // 组态非法（|fD|>1 或非有限系数，锁存） [-] / Illegal configuration, latched
    bError  : BOOL;           // 故障标志（与 bCfgBad 同源，R191 配对） [-] / Error flag, paired with bCfgBad
END_VAR
VAR
    _bCfgLatch: BOOL;         // 组态非法锁存位（解除沿 = bReset 上升沿） / Latched config fault, cleared by reset edge
    rtReset   : R_TRIG;       // 复位沿实例，段 0 无条件调用 / Reset edge instance
    _bNonFin  : BOOL;         // 输入非有限当拍量 [-] / Non-finite input this scan
    _fRaw1    : LREAL;        // 当拍回路 1 未钳解耦值 [%] / Unlimited decoupled value for loop 1
    _fRaw2    : LREAL;        // 当拍回路 2 未钳解耦值 [%] / Unlimited decoupled value for loop 2
END_VAR
VAR CONSTANT
    DL_DC2_UMIN : LREAL := 0.0;    // 输出行程下限 [%] / Output travel floor [%]
    DL_DC2_UMAX : LREAL := 100.0;  // 输出行程上限 [%] / Output travel ceiling [%]
    DL_DC2_ONE  : LREAL := 1.0;    // 系数域界（|fD| 上限） [无量纲] / Factor domain bound
    DL_DC2_EPS  : LREAL := 0.0;    // 非有限差值判零基准 [-] / Non-finite difference zero base
END_VAR

(* —— 段 0：非有限判 + 组态闸 + 沿刷新 —— *)
_bNonFin := (fU1 <> fU1) OR ((fU1 - fU1) <> DL_DC2_EPS)
         OR (fU2 <> fU2) OR ((fU2 - fU2) <> DL_DC2_EPS);        // 主控输出非有限（R245） / Non-finite controller outputs
IF (ABS(fD12) > DL_DC2_ONE) OR (ABS(fD21) > DL_DC2_ONE)
   OR (fD12 <> fD12) OR ((fD12 - fD12) <> DL_DC2_EPS)
   OR (fD21 <> fD21) OR ((fD21 - fD21) <> DL_DC2_EPS) THEN
    _bCfgLatch := TRUE;                                         // 系数越域/非有限：锁存（R188 解除沿 = bReset 上升沿） / Factor out of domain: latch
END_IF
rtReset(CLK := bReset);                                         // 复位沿，每拍必调 / Reset edge, every scan

(* —— 段 1：复位沿 —— *)
IF rtReset.Q THEN
    _bCfgLatch := FALSE;                                        // 清组态非法锁存 / Clear cfg latch
END_IF

(* —— 段 2：解耦主算（直通条件三支：未使能 / 组态非法 / 输出非有限） —— *)
IF (NOT bEnable) OR _bCfgLatch OR _bNonFin THEN
    fU1Eff := fU1;                                              // 直通：回路 1 原值（头注释②④声明） / Bypass loop 1
    fU2Eff := fU2;                                              // 直通：回路 2 原值 / Bypass loop 2
ELSE
    _fRaw1 := fU1 + fD21 * fU2;                                 // 静态解耦注入：u2 对回路 1 的影响补偿 / Static decoupling injection onto loop 1
    _fRaw2 := fU2 + fD12 * fU1;                                 // 静态解耦注入：u1 对回路 2 的影响补偿 / Static decoupling injection onto loop 2
    IF _fRaw1 > DL_DC2_UMAX THEN
        fU1Eff := DL_DC2_UMAX;                                  // 回路 1 上钳 100% / Clamp loop 1 high
    ELSIF _fRaw1 < DL_DC2_UMIN THEN
        fU1Eff := DL_DC2_UMIN;                                  // 回路 1 下钳 0% / Clamp loop 1 low
    ELSE
        fU1Eff := _fRaw1;                                       // 行程内接受 / In-travel accept
    END_IF
    IF _fRaw2 > DL_DC2_UMAX THEN
        fU2Eff := DL_DC2_UMAX;                                  // 回路 2 上钳 / Clamp loop 2 high
    ELSIF _fRaw2 < DL_DC2_UMIN THEN
        fU2Eff := DL_DC2_UMIN;                                  // 回路 2 下钳 / Clamp loop 2 low
    ELSE
        fU2Eff := _fRaw2;                                       // 行程内接受 / In-travel accept
    END_IF
END_IF

(* —— 段 3：出口单点映射（名实双出口同源，R191） —— *)
bEnabled := bEnable AND (NOT _bCfgLatch);                       // 生效指示 = 使能 ∧ 组态合法 / Active = enabled and config valid
bCfgBad  := _bCfgLatch;                                         // 组态非法出口 / Cfg fault outlet
bError   := _bCfgLatch;                                         // 故障标志与 bCfgBad 同源 / Error flag same source

END_FUNCTION_BLOCK

(* ---- FB_DL_DerivativeNoiseWeight.st ---- *)
(*
  Name        : FB_DL_DerivativeNoiseWeight
  Category    : DL_Algo
  Version     : 1.0.0
  Purpose     : 微分项噪声权重与降权：以原始微分为基准，用低通差分残差估计高频能量占比，占比超阈时按比例衰减有效微分增益 Kd，抑制噪声放大而不改 PidController 契约；/ Derivative noise weighting: estimate high-frequency energy share from the residual between raw and low-passed derivative, and attenuate the effective Kd proportionally when the share exceeds threshold
  溯源        : 借 t2-5-modpid·deriv 的分类/参数域组织，clean-room 实现
  Boundary    : ① 采样周期闸：tDt <= T#0S → 锁存故障（除零前置，dt 秒化后仍 > eps）；
                ② 能量比除子闸：eSig + eHf <= eps → 占比按 0 处理（不产生 Inf/NaN）；
                ③ 非有限输入该拍不推进差分与能量估计（保留上拍值，防污染 EMA）；
                ④ 衰减上限钳位 fAttenMax ∈ [0,1]，KdEff >= KdNom·(1-fAttenMax) 不会取负；
                ⑤ 本件只作观测器输出，不修改任何控制回路参数（属主边界声明）。
*)
TYPE E_DL_DnwState :
(
    eIdle  := 0,                             (* 未使能 / Disabled *)
    eRun   := 10,                            (* 观测运行 / Observing *)
    eFault := 90                             (* 故障锁存相 / Fault latched *)
);
END_TYPE

TYPE E_DL_DnwCause :
(
    eNone       := 0,                        (* 无故障成因 / No cause *)
    eCfgIllegal := 1,                        (* 组态非法：周期/增益/阈值越域 / Illegal config *)
    ePhaseBad   := 2                         (* 非法相位兜底 / Illegal phase fallback *)
);
END_TYPE

FUNCTION_BLOCK FB_DL_DerivativeNoiseWeight
VAR_INPUT
    fIn        : REAL := 0.0;                (* 反馈测量输入（PV）[工程单位] / Feedback measurement *)
    tDt        : TIME := T#10MS;             (* 采样周期（微分除子），域 > T#0S [ms] / Sampling period, must be > 0 *)
    fKdNom     : REAL := 1.0;                (* 标称微分增益（不动原参数），域 > 0 [s] / Nominal derivative gain, > 0 *)
    fRatioThr  : REAL := 0.3;                (* 高频能量占比阈值，域 (0,1) [-] / High-frequency ratio threshold *)
    fAttenMax  : REAL := 0.9;                (* 最大衰减比，域 [0,1] [-] / Maximum attenuation ratio *)
    fBeta      : REAL := 0.1;                (* 低通/能量 EMA 权重，域 (0,1] [-] / Filter and energy EMA weight *)
    bEnable    : BOOL := TRUE;               (* 使能 [-] / Enable *)
    bReset     : BOOL := FALSE;              (* 复位命令，上升沿清估计与输出 [-] / Reset command *)
END_VAR
VAR_OUTPUT
    fDerivRaw  : REAL;                       (* 原始微分（未滤波）[工程单位/s] / Raw derivative *)
    fDerivFilt : REAL;                       (* 低通微分 [工程单位/s] / Low-passed derivative *)
    fHfRatio   : REAL;                       (* 高频能量占比 0..1 [-] / High-frequency energy ratio *)
    fKdEff     : REAL;                       (* 降权后有效微分增益 [s] / Effective attenuated derivative gain *)
    bAtten     : BOOL;                       (* 降权生效指示 [-] / Attenuation active *)
    eState     : E_DL_DnwState;              (* 状态出口 / State outlet *)
    eCause     : E_DL_DnwCause;              (* 故障成因出口（R190 归因唯一） / Fault cause outlet *)
    bError     : BOOL;                       (* 故障锁存标志 [-] / Fault latch flag *)
END_VAR
VAR
    _eState  : E_DL_DnwState := E_DL_DnwState.eIdle;     (* 内部相位（CASE 唯一写入目标） / Internal phase *)
    _eCause  : E_DL_DnwCause := E_DL_DnwCause.eNone;     (* 故障成因锁存量 / Latched cause *)
    rtReset  : R_TRIG;                       (* 复位沿实例，段 0 无条件调用 / Reset edge instance *)
    _bFault  : BOOL;                         (* 故障锁存位 / Latched fault bit *)
    _bCfgBad : BOOL;                         (* 组态非法当拍量 / Illegal config this scan *)
    _bInit   : BOOL;                         (* 前值初始化标志（首拍不产虚假微分尖峰） / First-scan init *)
    _bFinite : BOOL;                         (* 输入有限性当拍量 / Input finiteness *)
    _fPrev   : REAL;                         (* 上拍输入快照 [工程单位] / Previous input *)
    _fDtSec  : REAL;                         (* 采样周期折算秒值，域 > eps [s] / Sampling period in seconds *)
    _fHf     : REAL;                         (* 高频残差 = 原始 - 低通 [工程单位/s] / High-frequency residual *)
    _fEHf    : REAL;                         (* 高频能量 EMA [工程单位²/s²] / High-frequency energy EMA *)
    _fESig   : REAL;                         (* 低通信号能量 EMA [工程单位²/s²] / Signal energy EMA *)
    _fRatio  : REAL;                         (* 未钳位占比 [-] / Unclamped ratio *)
    _fAtten  : REAL;                         (* 本拍衰减比 0..fAttenMax [-] / Attenuation this scan *)
END_VAR
VAR CONSTANT
    DL_DNW_EPS : REAL := 1.0E-6;             (* 判零容差（REAL 量级）[-] / Epsilon *)
    DL_DNW_ONE : REAL := 1.0;                (* 实数 1 常量 [-] / Real one *)
    DL_DNW_ZERO: REAL := 0.0;                (* 实数零常量 [-] / Real zero *)
END_VAR

(* —— 段 0：当拍判据派生 + 实例无条件刷新（R228A） —— *)
_fDtSec := TIME_TO_LREAL(tDt) / 1000.0;                                        (* 周期秒化（除子为常量 1000，无除零） / Period to seconds *)
_bCfgBad := NOT (tDt > T#0S)                                                   (* 周期正域闸（除零前置） / Period gate *)
            OR (fKdNom <= DL_DNW_EPS)                                          (* 微分增益正域闸 / Kd positive gate *)
            OR (fRatioThr <= DL_DNW_EPS) OR (fRatioThr >= DL_DNW_ONE)          (* 阈值域闸 (0,1) / Threshold gate *)
            OR (fAttenMax < DL_DNW_ZERO) OR (fAttenMax > DL_DNW_ONE)           (* 衰减比域闸 [0,1] / Attenuation gate *)
            OR (fBeta <= DL_DNW_EPS) OR (fBeta > DL_DNW_ONE);                  (* EMA 系数域闸 (0,1] / EMA weight gate *)
rtReset(CLK := bReset);                                                        (* 复位沿每拍必调 / Reset edge every scan *)
_bFinite := (fIn = fIn) AND ((fIn - fIn) = (fIn - fIn));                       (* NaN 自反 + Inf 差判联合闸 / NaN and Inf gate *)

(* —— 段 1：单拍量预清零（R107） —— *)
bAtten := FALSE;                                                               (* 降权指示预清 / Attenuation preset *)
_fAtten := DL_DNW_ZERO;                                                        (* 衰减比预清 / Attenuation preset *)

(* —— 段 2：复位沿处理（作用域：清故障 + 清估计 + 清初始化 + 迁 eIdle，R283 逐项声明） —— *)
IF rtReset.Q THEN
    _bFault := FALSE;                                                          (* 清故障锁存 / Clear fault *)
    _eCause := E_DL_DnwCause.eNone;                                            (* 清成因 / Clear cause *)
    _fPrev := DL_DNW_ZERO;                                                     (* 清前值 / Clear previous *)
    _fHf := DL_DNW_ZERO;                                                       (* 清高频残差 / Clear residual *)
    _fEHf := DL_DNW_ZERO;                                                      (* 清高频能量 / Clear hf energy *)
    _fESig := DL_DNW_ZERO;                                                     (* 清信号能量 / Clear signal energy *)
    _bInit := FALSE;                                                           (* 清初始化标志 / Clear init *)
    fDerivRaw := DL_DNW_ZERO;                                                  (* 清原始微分出口 / Clear raw outlet *)
    fDerivFilt := DL_DNW_ZERO;                                                 (* 清低通微分出口 / Clear filtered outlet *)
    fHfRatio := DL_DNW_ZERO;                                                   (* 清占比出口 / Clear ratio outlet *)
    fKdEff := fKdNom;                                                          (* 有效增益回标称（无降权基准） / Effective gain back to nominal *)
    _eState := E_DL_DnwState.eIdle;                                            (* 迁未使能相 / Back to idle *)
END_IF

(* —— 段 3：组态故障锁存（锁存至复位沿，R189） —— *)
IF _bCfgBad AND NOT _bFault THEN
    _bFault := TRUE;                                                           (* 锁存故障位 / Latch fault *)
    _eCause := E_DL_DnwCause.eCfgIllegal;                                      (* 成因：组态非法 / Cause: illegal config *)
    _eState := E_DL_DnwState.eFault;                                           (* 同步迁故障相 / Migrate to fault *)
END_IF

(* —— 段 4：CASE 主状态机（ELSE 兜底迁 eFault，红线 6） —— *)
CASE _eState OF
    E_DL_DnwState.eIdle:                                                       (* 未使能：输出回标称基准 / Disabled *)
        fKdEff := fKdNom;                                                      (* 无降权：有效增益 = 标称 / No attenuation *)
        _bInit := FALSE;                                                       (* 失能清初始化 / Clear init *)
        IF bEnable AND NOT _bFault THEN
            _eState := E_DL_DnwState.eRun;                                     (* 使能进入观测 / Enter observing *)
        END_IF
    E_DL_DnwState.eRun:                                                        (* 观测相：微分 + 能量分离 + 降权 / Observing *)
        IF NOT bEnable THEN
            _eState := E_DL_DnwState.eIdle;                                    (* 失能回未使能 / Back to idle *)
        ELSIF _bFinite AND (_fDtSec > DL_DNW_EPS) THEN
            IF NOT _bInit THEN
                _fPrev := fIn;                                                 (* 首拍对齐：防虚假微分尖峰 / First-scan alignment *)
                _bInit := TRUE;                                                (* 立初始化标志 / Set init *)
            END_IF
            fDerivRaw := (fIn - _fPrev) / _fDtSec;                             (* 原始微分：除子 dt 已过闸 > eps [工程单位/s] / Raw derivative, divisor gated *)
            fDerivFilt := fDerivFilt + fBeta * (fDerivRaw - fDerivFilt);       (* 一阶低通（EMA 形式，系数 (0,1]） / First-order low pass *)
            _fHf := fDerivRaw - fDerivFilt;                                    (* 高频残差：低通漏掉的快变成分 / High-frequency residual *)
            _fEHf := (1.0 - fBeta) * _fEHf + fBeta * _fHf * _fHf;              (* 高频能量 EMA（平方项恒非负） / HF energy EMA *)
            _fESig := (1.0 - fBeta) * _fESig + fBeta * fDerivFilt * fDerivFilt; (* 信号能量 EMA / Signal energy EMA *)
            _fPrev := fIn;                                                     (* 前值推进（仅有限拍推进） / Advance previous *)
            IF (_fEHf + _fESig) > DL_DNW_EPS THEN
                _fRatio := _fEHf / (_fEHf + _fESig);                           (* 占比：除子已过闸（边界②） / Ratio, divisor gated *)
            ELSE
                _fRatio := DL_DNW_ZERO;                                        (* 能量全零：占比按 0（无噪声语义） / Zero energy: ratio 0 *)
            END_IF
            IF _fRatio < DL_DNW_ZERO THEN
                _fRatio := DL_DNW_ZERO;                                        (* 下限兜底（数值噪声防负） / Lower fallback *)
            ELSIF _fRatio > DL_DNW_ONE THEN
                _fRatio := DL_DNW_ONE;                                         (* 上限饱和 1.0 / Upper saturation *)
            END_IF
            fHfRatio := _fRatio;                                               (* 占比出口 / Ratio outlet *)
            IF _fRatio > fRatioThr THEN
                _fAtten := fAttenMax * (_fRatio - fRatioThr) / (1.0 - fRatioThr);   (* 超阈后线性升权衰减（除子 < 1 且已过闸） / Linear attenuation beyond threshold *)
                IF _fAtten > fAttenMax THEN
                    _fAtten := fAttenMax;                                      (* 衰减上限钳位 / Attenuation cap *)
                ELSIF _fAtten < DL_DNW_ZERO THEN
                    _fAtten := DL_DNW_ZERO;                                    (* 衰减下限钳位 / Attenuation floor *)
                END_IF
                bAtten := TRUE;                                                (* 降权生效 / Attenuation active *)
            END_IF
            fKdEff := fKdNom * (1.0 - _fAtten);                                (* 有效增益：_fAtten <= 1 保证非负（边界④） / Effective gain, non-negative *)
        END_IF                                                                 (* 非有限输入：全部估计保持上拍（边界③） / Non-finite: hold *)
    E_DL_DnwState.eFault:                                                      (* 故障相：冻结保持末值，仅复位沿出 / Fault *)
        ;                                                                      (* 锁存回放（R28） / Replay from latch *)
    ELSE                                                                       (* 非法相位兜底迁安全态 / Illegal phase fallback *)
        _eState := E_DL_DnwState.eFault;                                       (* 迁故障相 / To fault *)
        _bFault := TRUE;                                                       (* 同步锁存 / Latch *)
        _eCause := E_DL_DnwCause.ePhaseBad;                                    (* 成因：非法相位 / Cause: illegal phase *)
END_CASE

(* —— 段 5：出口映射（bError/eState 同源，R191） —— *)
bError := _bFault;                                                             (* 故障标志镜像 / Fault flag mirror *)
eState := _eState;                                                             (* 状态出口 / State outlet *)
eCause := _eCause;                                                             (* 成因出口 / Cause outlet *)
END_FUNCTION_BLOCK
